  movel([0.274819, -1.341479, -2.579880, -0.791030, 1.570796, 1.845616],accel_mss,speed_ms,0,blend_radius_m)
  movel([0.275794, -1.341271, -2.580017, -0.791101, 1.570796, 1.846590],accel_mss,speed_ms,0,blend_radius_m)
  movel([0.276766, -1.341079, -2.580143, -0.791167, 1.570796, 1.847563],accel_mss,speed_ms,0,blend_radius_m)
  movel([0.277679, -1.340913, -2.580252, -0.791224, 1.570796, 1.848475],accel_mss,speed_ms,0,blend_radius_m)
  movel([0.278587, -1.340762, -2.580351, -0.791276, 1.570796, 1.849384],accel_mss,speed_ms,0,blend_radius_m)
  movel([0.278988, -1.340706, -2.580387, -0.791295, 1.570796, 1.849784],accel_mss,speed_ms,0,blend_radius_m)
  movel([0.279382, -1.340663, -2.580416, -0.791310, 1.570796, 1.850178],accel_mss,speed_ms,0,blend_radius_m)
  movel([0.279771, -1.340637, -2.580433, -0.791319, 1.570796, 1.850568],accel_mss,speed_ms,0,blend_radius_m)
  movel([0.279984, -1.340628, -2.580439, -0.791322, 1.570796, 1.850780],accel_mss,speed_ms,0,blend_radius_m)
  movel([0.280191, -1.340629, -2.580438, -0.791322, 1.570796, 1.850987],accel_mss,speed_ms,0,blend_radius_m)
  movel([0.280203, -1.340637, -2.580433, -0.791319, 1.570796, 1.850999],accel_mss,speed_ms,0,blend_radius_m)
  movel([0.280197, -1.340656, -2.580421, -0.791313, 1.570796, 1.850993],accel_mss,speed_ms,0,blend_radius_m)
  movel([0.280179, -1.340667, -2.580413, -0.791309, 1.570796, 1.850976],accel_mss,speed_ms,0,blend_radius_m)
  speed_ms = 0.003
  movel([0.280179, -1.327920, -2.574072, -0.810397, 1.570796, 1.850976],accel_mss,speed_ms,0,blend_radius_m)
  speed_ms = 0.01
  movel([0.280179, -1.303552, -2.561012, -0.847825, 1.570796, 1.850976],accel_mss,speed_ms,0,blend_radius_m)
  movel([0.262380, -1.358037, -2.525199, -0.829153, 1.570796, 1.833176],accel_mss,speed_ms,0,blend_radius_m)
  movel([0.262380, -1.381577, -2.537576, -0.793236, 1.570796, 1.833176],accel_mss,speed_ms,0,blend_radius_m)
  speed_ms = 0.003
  movel([0.262380, -1.390744, -2.542086, -0.779559, 1.570796, 1.833176],accel_mss,speed_ms,0,blend_radius_m)
  speed_ms = 0.007
  movel([0.261890, -1.392448, -2.540846, -0.779096, 1.570796, 1.832686],accel_mss,speed_ms,0,blend_radius_m)
  movel([0.261638, -1.393307, -2.540218, -0.778864, 1.570796, 1.832434],accel_mss,speed_ms,0,blend_radius_m)
  movel([0.261560, -1.393546, -2.540044, -0.778799, 1.570796, 1.832357],accel_mss,speed_ms,0,blend_radius_m)
  movel([0.261476, -1.393785, -2.539869, -0.778735, 1.570796, 1.832272],accel_mss,speed_ms,0,blend_radius_m)
  movel([0.261419, -1.393927, -2.539765, -0.778697, 1.570796, 1.832216],accel_mss,speed_ms,0,blend_radius_m)
  movel([0.261357, -1.394067, -2.539663, -0.778659, 1.570796, 1.832153],accel_mss,speed_ms,0,blend_radius_m)
  movel([0.261341, -1.394090, -2.539646, -0.778653, 1.570796, 1.832137],accel_mss,speed_ms,0,blend_radius_m)
  movel([0.261318, -1.394107, -2.539633, -0.778648, 1.570796, 1.832114],accel_mss,speed_ms,0,blend_radius_m)
  movel([0.261293, -1.394115, -2.539628, -0.778646, 1.570796, 1.832090],accel_mss,speed_ms,0,blend_radius_m)
  movel([0.261271, -1.394116, -2.539627, -0.778646, 1.570796, 1.832067],accel_mss,speed_ms,0,blend_radius_m)
  movel([0.256001, -1.393339, -2.540195, -0.778855, 1.570796, 1.826797],accel_mss,speed_ms,0,blend_radius_m)
  movel([0.256257, -1.392428, -2.540860, -0.779101, 1.570796, 1.827054],accel_mss,speed_ms,0,blend_radius_m)
  movel([0.256515, -1.391516, -2.541524, -0.779349, 1.570796, 1.827311],accel_mss,speed_ms,0,blend_radius_m)
  movel([0.259448, -1.391126, -2.541808, -0.779455, 1.570796, 1.830244],accel_mss,speed_ms,0,blend_radius_m)
  movel([0.262380, -1.390744, -2.542086, -0.779559, 1.570796, 1.833176],accel_mss,speed_ms,0,blend_radius_m)
  speed_ms = 0.003
  movel([0.262380, -1.393840, -2.543573, -0.774975, 1.570796, 1.833176],accel_mss,speed_ms,0,blend_radius_m)
  speed_ms = 0.007
  movel([0.261890, -1.395540, -2.542330, -0.774519, 1.570796, 1.832686],accel_mss,speed_ms,0,blend_radius_m)
  movel([0.261638, -1.396398, -2.541701, -0.774290, 1.570796, 1.832434],accel_mss,speed_ms,0,blend_radius_m)
  movel([0.261560, -1.396636, -2.541527, -0.774227, 1.570796, 1.832357],accel_mss,speed_ms,0,blend_radius_m)
  movel([0.261476, -1.396875, -2.541351, -0.774163, 1.570796, 1.832272],accel_mss,speed_ms,0,blend_radius_m)
  movel([0.261419, -1.397016, -2.541248, -0.774126, 1.570796, 1.832216],accel_mss,speed_ms,0,blend_radius_m)
  movel([0.261357, -1.397155, -2.541145, -0.774089, 1.570796, 1.832153],accel_mss,speed_ms,0,blend_radius_m)
  movel([0.261341, -1.397178, -2.541128, -0.774083, 1.570796, 1.832137],accel_mss,speed_ms,0,blend_radius_m)
  movel([0.261318, -1.397196, -2.541115, -0.774078, 1.570796, 1.832114],accel_mss,speed_ms,0,blend_radius_m)
  movel([0.261293, -1.397203, -2.541110, -0.774076, 1.570796, 1.832090],accel_mss,speed_ms,0,blend_radius_m)
  movel([0.261271, -1.397204, -2.541109, -0.774076, 1.570796, 1.832067],accel_mss,speed_ms,0,blend_radius_m)
  movel([0.256001, -1.396429, -2.541678, -0.774282, 1.570796, 1.826797],accel_mss,speed_ms,0,blend_radius_m)
  movel([0.256257, -1.395521, -2.542344, -0.774524, 1.570796, 1.827054],accel_mss,speed_ms,0,blend_radius_m)
  movel([0.256515, -1.394611, -2.543010, -0.774768, 1.570796, 1.827311],accel_mss,speed_ms,0,blend_radius_m)
  movel([0.259448, -1.394222, -2.543295, -0.774872, 1.570796, 1.830244],accel_mss,speed_ms,0,blend_radius_m)
  movel([0.262380, -1.393840, -2.543573, -0.774975, 1.570796, 1.833176],accel_mss,speed_ms,0,blend_radius_m)
  speed_ms = 0.003
  movel([0.262380, -1.381577, -2.537576, -0.793236, 1.570796, 1.833176],accel_mss,speed_ms,0,blend_radius_m)
  speed_ms = 0.01
  movel([0.262380, -1.358037, -2.525199, -0.829153, 1.570796, 1.833176],accel_mss,speed_ms,0,blend_radius_m)
  movel([0.278975, -1.298309, -2.564258, -0.849822, 1.570796, 1.849771],accel_mss,speed_ms,0,blend_radius_m)
  movel([0.278975, -1.322751, -2.577384, -0.812254, 1.570796, 1.849771],accel_mss,speed_ms,0,blend_radius_m)
  speed_ms = 0.003
  movel([0.278975, -1.332307, -2.582178, -0.797904, 1.570796, 1.849771],accel_mss,speed_ms,0,blend_radius_m)
  speed_ms = 0.007
  movel([0.275846, -1.332753, -2.581889, -0.797747, 1.570796, 1.846643],accel_mss,speed_ms,0,blend_radius_m)
  movel([0.272717, -1.333207, -2.581595, -0.797586, 1.570796, 1.843513],accel_mss,speed_ms,0,blend_radius_m)
  movel([0.273170, -1.331664, -2.582593, -0.798132, 1.570796, 1.843966],accel_mss,speed_ms,0,blend_radius_m)
  movel([0.273625, -1.330114, -2.583591, -0.798683, 1.570796, 1.844422],accel_mss,speed_ms,0,blend_radius_m)
  movel([0.274406, -1.330222, -2.583522, -0.798645, 1.570796, 1.845202],accel_mss,speed_ms,0,blend_radius_m)
  movel([0.274838, -1.330281, -2.583484, -0.798624, 1.570796, 1.845634],accel_mss,speed_ms,0,blend_radius_m)
  movel([0.275574, -1.330385, -2.583417, -0.798587, 1.570796, 1.846370],accel_mss,speed_ms,0,blend_radius_m)
  movel([0.276428, -1.330502, -2.583342, -0.798545, 1.570796, 1.847224],accel_mss,speed_ms,0,blend_radius_m)
  movel([0.277289, -1.330626, -2.583262, -0.798501, 1.570796, 1.848086],accel_mss,speed_ms,0,blend_radius_m)
  movel([0.279389, -1.330926, -2.583069, -0.798394, 1.570796, 1.850186],accel_mss,speed_ms,0,blend_radius_m)
  movel([0.279182, -1.331618, -2.582623, -0.798149, 1.570796, 1.849978],accel_mss,speed_ms,0,blend_radius_m)
  movel([0.278975, -1.332307, -2.582178, -0.797904, 1.570796, 1.849771],accel_mss,speed_ms,0,blend_radius_m)
  speed_ms = 0.003
  movel([0.278975, -1.335541, -2.583759, -0.793089, 1.570796, 1.849771],accel_mss,speed_ms,0,blend_radius_m)
  speed_ms = 0.007
  movel([0.275846, -1.335986, -2.583470, -0.792933, 1.570796, 1.846643],accel_mss,speed_ms,0,blend_radius_m)
  movel([0.272717, -1.336439, -2.583175, -0.792775, 1.570796, 1.843513],accel_mss,speed_ms,0,blend_radius_m)
  movel([0.273170, -1.334899, -2.584176, -0.793315, 1.570796, 1.843966],accel_mss,speed_ms,0,blend_radius_m)
  movel([0.273625, -1.333353, -2.585176, -0.793860, 1.570796, 1.844422],accel_mss,speed_ms,0,blend_radius_m)
  movel([0.274406, -1.333460, -2.585107, -0.793822, 1.570796, 1.845202],accel_mss,speed_ms,0,blend_radius_m)
  movel([0.274838, -1.333519, -2.585069, -0.793801, 1.570796, 1.845634],accel_mss,speed_ms,0,blend_radius_m)
  movel([0.275574, -1.333622, -2.585002, -0.793765, 1.570796, 1.846370],accel_mss,speed_ms,0,blend_radius_m)
  movel([0.276428, -1.333739, -2.584926, -0.793723, 1.570796, 1.847224],accel_mss,speed_ms,0,blend_radius_m)
  movel([0.277289, -1.333863, -2.584846, -0.793680, 1.570796, 1.848086],accel_mss,speed_ms,0,blend_radius_m)
  movel([0.279389, -1.334162, -2.584653, -0.793574, 1.570796, 1.850186],accel_mss,speed_ms,0,blend_radius_m)
  movel([0.279182, -1.334853, -2.584205, -0.793331, 1.570796, 1.849978],accel_mss,speed_ms,0,blend_radius_m)
  movel([0.278975, -1.335541, -2.583759, -0.793089, 1.570796, 1.849771],accel_mss,speed_ms,0,blend_radius_m)
  speed_ms = 0.003
  movel([0.278975, -1.322751, -2.577384, -0.812254, 1.570796, 1.849771],accel_mss,speed_ms,0,blend_radius_m)
  speed_ms = 0.01
  movel([0.278975, -1.298309, -2.564258, -0.849822, 1.570796, 1.849771],accel_mss,speed_ms,0,blend_radius_m)
  movel([0.264711, -1.307973, -2.558248, -0.846168, 1.570796, 1.835507],accel_mss,speed_ms,0,blend_radius_m)
  movel([0.264711, -1.332279, -2.571252, -0.808858, 1.570796, 1.835507],accel_mss,speed_ms,0,blend_radius_m)
  speed_ms = 0.003
  movel([0.264711, -1.341777, -2.575999, -0.794614, 1.570796, 1.835507],accel_mss,speed_ms,0,blend_radius_m)
  speed_ms = 0.007
  movel([0.264715, -1.341787, -2.575992, -0.794610, 1.570796, 1.835511],accel_mss,speed_ms,0,blend_radius_m)
  movel([0.264709, -1.341799, -2.575984, -0.794606, 1.570796, 1.835505],accel_mss,speed_ms,0,blend_radius_m)
  movel([0.264688, -1.341820, -2.575970, -0.794599, 1.570796, 1.835485],accel_mss,speed_ms,0,blend_radius_m)
  movel([0.264666, -1.341839, -2.575957, -0.794592, 1.570796, 1.835463],accel_mss,speed_ms,0,blend_radius_m)
  movel([0.264589, -1.341894, -2.575921, -0.794574, 1.570796, 1.835385],accel_mss,speed_ms,0,blend_radius_m)
  movel([0.264497, -1.341950, -2.575884, -0.794555, 1.570796, 1.835293],accel_mss,speed_ms,0,blend_radius_m)
  movel([0.264400, -1.341999, -2.575852, -0.794538, 1.570796, 1.835196],accel_mss,speed_ms,0,blend_radius_m)
  movel([0.264310, -1.342037, -2.575827, -0.794525, 1.570796, 1.835107],accel_mss,speed_ms,0,blend_radius_m)
  movel([0.264246, -1.342053, -2.575816, -0.794520, 1.570796, 1.835043],accel_mss,speed_ms,0,blend_radius_m)
  movel([0.264232, -1.342053, -2.575816, -0.794520, 1.570796, 1.835028],accel_mss,speed_ms,0,blend_radius_m)
  movel([0.264222, -1.342048, -2.575820, -0.794521, 1.570796, 1.835018],accel_mss,speed_ms,0,blend_radius_m)
  movel([0.264217, -1.342037, -2.575827, -0.794525, 1.570796, 1.835014],accel_mss,speed_ms,0,blend_radius_m)
  movel([0.264223, -1.342025, -2.575835, -0.794529, 1.570796, 1.835020],accel_mss,speed_ms,0,blend_radius_m)
  movel([0.264244, -1.342004, -2.575849, -0.794536, 1.570796, 1.835040],accel_mss,speed_ms,0,blend_radius_m)
  movel([0.264266, -1.341985, -2.575861, -0.794543, 1.570796, 1.835062],accel_mss,speed_ms,0,blend_radius_m)
  movel([0.264341, -1.341931, -2.575897, -0.794561, 1.570796, 1.835137],accel_mss,speed_ms,0,blend_radius_m)
  movel([0.264435, -1.341874, -2.575934, -0.794581, 1.570796, 1.835232],accel_mss,speed_ms,0,blend_radius_m)
  movel([0.264532, -1.341826, -2.575966, -0.794597, 1.570796, 1.835329],accel_mss,speed_ms,0,blend_radius_m)
  movel([0.264622, -1.341788, -2.575991, -0.794610, 1.570796, 1.835418],accel_mss,speed_ms,0,blend_radius_m)
  movel([0.264683, -1.341772, -2.576002, -0.794616, 1.570796, 1.835480],accel_mss,speed_ms,0,blend_radius_m)
  movel([0.264700, -1.341771, -2.576002, -0.794616, 1.570796, 1.835496],accel_mss,speed_ms,0,blend_radius_m)
  movel([0.264711, -1.341777, -2.575999, -0.794614, 1.570796, 1.835507],accel_mss,speed_ms,0,blend_radius_m)
  speed_ms = 0.003
  movel([0.264711, -1.344989, -2.577565, -0.789835, 1.570796, 1.835507],accel_mss,speed_ms,0,blend_radius_m)
  speed_ms = 0.007
  movel([0.264715, -1.345000, -2.577558, -0.789832, 1.570796, 1.835511],accel_mss,speed_ms,0,blend_radius_m)
  movel([0.264709, -1.345012, -2.577550, -0.789827, 1.570796, 1.835505],accel_mss,speed_ms,0,blend_radius_m)
  movel([0.264688, -1.345033, -2.577536, -0.789820, 1.570796, 1.835485],accel_mss,speed_ms,0,blend_radius_m)
  movel([0.264666, -1.345052, -2.577523, -0.789814, 1.570796, 1.835463],accel_mss,speed_ms,0,blend_radius_m)
  movel([0.264589, -1.345106, -2.577487, -0.789796, 1.570796, 1.835385],accel_mss,speed_ms,0,blend_radius_m)
  movel([0.264497, -1.345163, -2.577450, -0.789777, 1.570796, 1.835293],accel_mss,speed_ms,0,blend_radius_m)
  movel([0.264400, -1.345211, -2.577418, -0.789760, 1.570796, 1.835196],accel_mss,speed_ms,0,blend_radius_m)
  movel([0.264310, -1.345249, -2.577393, -0.789747, 1.570796, 1.835107],accel_mss,speed_ms,0,blend_radius_m)
  movel([0.264246, -1.345265, -2.577382, -0.789742, 1.570796, 1.835043],accel_mss,speed_ms,0,blend_radius_m)
  movel([0.264232, -1.345265, -2.577382, -0.789742, 1.570796, 1.835028],accel_mss,speed_ms,0,blend_radius_m)
  movel([0.264222, -1.345260, -2.577385, -0.789744, 1.570796, 1.835018],accel_mss,speed_ms,0,blend_radius_m)
  movel([0.264217, -1.345249, -2.577392, -0.789747, 1.570796, 1.835014],accel_mss,speed_ms,0,blend_radius_m)
  movel([0.264223, -1.345237, -2.577400, -0.789751, 1.570796, 1.835020],accel_mss,speed_ms,0,blend_radius_m)
  movel([0.264244, -1.345216, -2.577414, -0.789758, 1.570796, 1.835040],accel_mss,speed_ms,0,blend_radius_m)
  movel([0.264266, -1.345197, -2.577427, -0.789765, 1.570796, 1.835062],accel_mss,speed_ms,0,blend_radius_m)
  movel([0.264341, -1.345143, -2.577463, -0.789783, 1.570796, 1.835137],accel_mss,speed_ms,0,blend_radius_m)
  movel([0.264435, -1.345086, -2.577500, -0.789802, 1.570796, 1.835232],accel_mss,speed_ms,0,blend_radius_m)
  movel([0.264532, -1.345038, -2.577532, -0.789819, 1.570796, 1.835329],accel_mss,speed_ms,0,blend_radius_m)
  movel([0.264622, -1.345000, -2.577557, -0.789831, 1.570796, 1.835418],accel_mss,speed_ms,0,blend_radius_m)
  movel([0.264683, -1.344984, -2.577568, -0.789837, 1.570796, 1.835480],accel_mss,speed_ms,0,blend_radius_m)
  movel([0.264700, -1.344984, -2.577568, -0.789837, 1.570796, 1.835496],accel_mss,speed_ms,0,blend_radius_m)
  movel([0.264711, -1.344989, -2.577565, -0.789835, 1.570796, 1.835507],accel_mss,speed_ms,0,blend_radius_m)
  speed_ms = 0.003
  movel([0.264711, -1.332279, -2.571252, -0.808858, 1.570796, 1.835507],accel_mss,speed_ms,0,blend_radius_m)
  speed_ms = 0.01
  movel([0.264711, -1.307973, -2.558248, -0.846168, 1.570796, 1.835507],accel_mss,speed_ms,0,blend_radius_m)
  movel([0.264022, -1.308308, -2.558037, -0.846043, 1.570796, 1.834819],accel_mss,speed_ms,0,blend_radius_m)
  movel([0.264022, -1.332610, -2.571037, -0.808742, 1.570796, 1.834819],accel_mss,speed_ms,0,blend_radius_m)
  speed_ms = 0.003
  movel([0.264022, -1.342105, -2.575782, -0.794502, 1.570796, 1.834819],accel_mss,speed_ms,0,blend_radius_m)
  speed_ms = 0.007
  movel([0.264026, -1.342115, -2.575775, -0.794498, 1.570796, 1.834823],accel_mss,speed_ms,0,blend_radius_m)
  movel([0.264020, -1.342128, -2.575767, -0.794494, 1.570796, 1.834817],accel_mss,speed_ms,0,blend_radius_m)
  movel([0.264000, -1.342149, -2.575753, -0.794487, 1.570796, 1.834797],accel_mss,speed_ms,0,blend_radius_m)
  movel([0.263978, -1.342168, -2.575741, -0.794481, 1.570796, 1.834774],accel_mss,speed_ms,0,blend_radius_m)
  movel([0.263901, -1.342222, -2.575705, -0.794462, 1.570796, 1.834697],accel_mss,speed_ms,0,blend_radius_m)
  movel([0.263809, -1.342279, -2.575668, -0.794443, 1.570796, 1.834605],accel_mss,speed_ms,0,blend_radius_m)
  movel([0.263712, -1.342327, -2.575636, -0.794426, 1.570796, 1.834508],accel_mss,speed_ms,0,blend_radius_m)
  movel([0.263622, -1.342365, -2.575610, -0.794413, 1.570796, 1.834419],accel_mss,speed_ms,0,blend_radius_m)
  movel([0.263558, -1.342382, -2.575600, -0.794408, 1.570796, 1.834354],accel_mss,speed_ms,0,blend_radius_m)
  movel([0.263544, -1.342381, -2.575600, -0.794408, 1.570796, 1.834340],accel_mss,speed_ms,0,blend_radius_m)
  movel([0.263534, -1.342376, -2.575603, -0.794410, 1.570796, 1.834330],accel_mss,speed_ms,0,blend_radius_m)
  movel([0.263529, -1.342366, -2.575610, -0.794413, 1.570796, 1.834326],accel_mss,speed_ms,0,blend_radius_m)
  movel([0.263535, -1.342354, -2.575618, -0.794417, 1.570796, 1.834332],accel_mss,speed_ms,0,blend_radius_m)
  movel([0.263555, -1.342332, -2.575632, -0.794424, 1.570796, 1.834352],accel_mss,speed_ms,0,blend_radius_m)
  movel([0.263578, -1.342313, -2.575645, -0.794431, 1.570796, 1.834374],accel_mss,speed_ms,0,blend_radius_m)
  movel([0.263652, -1.342259, -2.575680, -0.794449, 1.570796, 1.834449],accel_mss,speed_ms,0,blend_radius_m)
  movel([0.263747, -1.342202, -2.575718, -0.794469, 1.570796, 1.834543],accel_mss,speed_ms,0,blend_radius_m)
  movel([0.263844, -1.342154, -2.575750, -0.794485, 1.570796, 1.834640],accel_mss,speed_ms,0,blend_radius_m)
  movel([0.263933, -1.342116, -2.575775, -0.794498, 1.570796, 1.834730],accel_mss,speed_ms,0,blend_radius_m)
  movel([0.263995, -1.342100, -2.575785, -0.794504, 1.570796, 1.834791],accel_mss,speed_ms,0,blend_radius_m)
  movel([0.264012, -1.342100, -2.575786, -0.794504, 1.570796, 1.834808],accel_mss,speed_ms,0,blend_radius_m)
  movel([0.264022, -1.342105, -2.575782, -0.794502, 1.570796, 1.834819],accel_mss,speed_ms,0,blend_radius_m)
  speed_ms = 0.003
  movel([0.264022, -1.345317, -2.577348, -0.789725, 1.570796, 1.834819],accel_mss,speed_ms,0,blend_radius_m)
  speed_ms = 0.007
  movel([0.264026, -1.345327, -2.577341, -0.789721, 1.570796, 1.834823],accel_mss,speed_ms,0,blend_radius_m)
  movel([0.264020, -1.345339, -2.577333, -0.789717, 1.570796, 1.834817],accel_mss,speed_ms,0,blend_radius_m)
  movel([0.264000, -1.345360, -2.577319, -0.789710, 1.570796, 1.834797],accel_mss,speed_ms,0,blend_radius_m)
  movel([0.263978, -1.345379, -2.577306, -0.789703, 1.570796, 1.834774],accel_mss,speed_ms,0,blend_radius_m)
  movel([0.263901, -1.345434, -2.577270, -0.789685, 1.570796, 1.834697],accel_mss,speed_ms,0,blend_radius_m)
  movel([0.263809, -1.345490, -2.577233, -0.789666, 1.570796, 1.834605],accel_mss,speed_ms,0,blend_radius_m)
  movel([0.263712, -1.345538, -2.577201, -0.789650, 1.570796, 1.834508],accel_mss,speed_ms,0,blend_radius_m)
  movel([0.263622, -1.345576, -2.577176, -0.789637, 1.570796, 1.834419],accel_mss,speed_ms,0,blend_radius_m)
  movel([0.263558, -1.345593, -2.577165, -0.789631, 1.570796, 1.834354],accel_mss,speed_ms,0,blend_radius_m)
  movel([0.263544, -1.345593, -2.577165, -0.789631, 1.570796, 1.834340],accel_mss,speed_ms,0,blend_radius_m)
  movel([0.263534, -1.345588, -2.577168, -0.789633, 1.570796, 1.834330],accel_mss,speed_ms,0,blend_radius_m)
  movel([0.263529, -1.345577, -2.577175, -0.789637, 1.570796, 1.834326],accel_mss,speed_ms,0,blend_radius_m)
  movel([0.263535, -1.345565, -2.577183, -0.789641, 1.570796, 1.834332],accel_mss,speed_ms,0,blend_radius_m)
  movel([0.263555, -1.345544, -2.577197, -0.789648, 1.570796, 1.834352],accel_mss,speed_ms,0,blend_radius_m)
  movel([0.263578, -1.345525, -2.577210, -0.789654, 1.570796, 1.834374],accel_mss,speed_ms,0,blend_radius_m)
  movel([0.263652, -1.345471, -2.577246, -0.789672, 1.570796, 1.834449],accel_mss,speed_ms,0,blend_radius_m)
  movel([0.263747, -1.345414, -2.577283, -0.789692, 1.570796, 1.834543],accel_mss,speed_ms,0,blend_radius_m)
  movel([0.263844, -1.345366, -2.577315, -0.789708, 1.570796, 1.834640],accel_mss,speed_ms,0,blend_radius_m)
  movel([0.263933, -1.345328, -2.577340, -0.789721, 1.570796, 1.834730],accel_mss,speed_ms,0,blend_radius_m)
  movel([0.263995, -1.345312, -2.577351, -0.789726, 1.570796, 1.834791],accel_mss,speed_ms,0,blend_radius_m)
  movel([0.264012, -1.345311, -2.577351, -0.789726, 1.570796, 1.834808],accel_mss,speed_ms,0,blend_radius_m)
  movel([0.264022, -1.345317, -2.577348, -0.789725, 1.570796, 1.834819],accel_mss,speed_ms,0,blend_radius_m)
  speed_ms = 0.003
  movel([0.264022, -1.332610, -2.571037, -0.808742, 1.570796, 1.834819],accel_mss,speed_ms,0,blend_radius_m)
  speed_ms = 0.01
  movel([0.264022, -1.308308, -2.558037, -0.846043, 1.570796, 1.834819],accel_mss,speed_ms,0,blend_radius_m)
  movel([0.248737, -1.294338, -2.566693, -0.851357, 1.570796, 1.819533],accel_mss,speed_ms,0,blend_radius_m)
  movel([0.248737, -1.318834, -2.579871, -0.813685, 1.570796, 1.819533],accel_mss,speed_ms,0,blend_radius_m)
  speed_ms = 0.003
  movel([0.248737, -1.328414, -2.584683, -0.799292, 1.570796, 1.819533],accel_mss,speed_ms,0,blend_radius_m)
  speed_ms = 0.007
  movel([0.248697, -1.328446, -2.584662, -0.799280, 1.570796, 1.819493],accel_mss,speed_ms,0,blend_radius_m)
  movel([0.248652, -1.328468, -2.584649, -0.799273, 1.570796, 1.819448],accel_mss,speed_ms,0,blend_radius_m)
  movel([0.245500, -1.329570, -2.583941, -0.798878, 1.570796, 1.816296],accel_mss,speed_ms,0,blend_radius_m)
  movel([0.242434, -1.330648, -2.583248, -0.798493, 1.570796, 1.813230],accel_mss,speed_ms,0,blend_radius_m)
  movel([0.242300, -1.330689, -2.583221, -0.798479, 1.570796, 1.813096],accel_mss,speed_ms,0,blend_radius_m)
  movel([0.242169, -1.330719, -2.583202, -0.798468, 1.570796, 1.812965],accel_mss,speed_ms,0,blend_radius_m)
  movel([0.242113, -1.330722, -2.583200, -0.798467, 1.570796, 1.812909],accel_mss,speed_ms,0,blend_radius_m)
  movel([0.242059, -1.330716, -2.583204, -0.798469, 1.570796, 1.812855],accel_mss,speed_ms,0,blend_radius_m)
  movel([0.240657, -1.330365, -2.583430, -0.798594, 1.570796, 1.811454],accel_mss,speed_ms,0,blend_radius_m)
  movel([0.239079, -1.329963, -2.583689, -0.798737, 1.570796, 1.809875],accel_mss,speed_ms,0,blend_radius_m)
  movel([0.237230, -1.329485, -2.583996, -0.798908, 1.570796, 1.808027],accel_mss,speed_ms,0,blend_radius_m)
  movel([0.231703, -1.328086, -2.584894, -0.799410, 1.570796, 1.802500],accel_mss,speed_ms,0,blend_radius_m)
  movel([0.232587, -1.326228, -2.586081, -0.800080, 1.570796, 1.803383],accel_mss,speed_ms,0,blend_radius_m)
  movel([0.232933, -1.325504, -2.586543, -0.800342, 1.570796, 1.803729],accel_mss,speed_ms,0,blend_radius_m)
  movel([0.233237, -1.324867, -2.586949, -0.800574, 1.570796, 1.804034],accel_mss,speed_ms,0,blend_radius_m)
  movel([0.233502, -1.324323, -2.587294, -0.800772, 1.570796, 1.804298],accel_mss,speed_ms,0,blend_radius_m)
  movel([0.233562, -1.324211, -2.587365, -0.800812, 1.570796, 1.804358],accel_mss,speed_ms,0,blend_radius_m)
  movel([0.233589, -1.324181, -2.587385, -0.800823, 1.570796, 1.804385],accel_mss,speed_ms,0,blend_radius_m)
  movel([0.233622, -1.324163, -2.587396, -0.800830, 1.570796, 1.804419],accel_mss,speed_ms,0,blend_radius_m)
  movel([0.233654, -1.324164, -2.587395, -0.800829, 1.570796, 1.804450],accel_mss,speed_ms,0,blend_radius_m)
  movel([0.234609, -1.324536, -2.587159, -0.800694, 1.570796, 1.805405],accel_mss,speed_ms,0,blend_radius_m)
  movel([0.235192, -1.324772, -2.587009, -0.800608, 1.570796, 1.805988],accel_mss,speed_ms,0,blend_radius_m)
  movel([0.235770, -1.325013, -2.586855, -0.800520, 1.570796, 1.806567],accel_mss,speed_ms,0,blend_radius_m)
  movel([0.236518, -1.325343, -2.586646, -0.800401, 1.570796, 1.807314],accel_mss,speed_ms,0,blend_radius_m)
  movel([0.237265, -1.325673, -2.586435, -0.800281, 1.570796, 1.808061],accel_mss,speed_ms,0,blend_radius_m)
  movel([0.239935, -1.326833, -2.585695, -0.799861, 1.570796, 1.810731],accel_mss,speed_ms,0,blend_radius_m)
  movel([0.240884, -1.327196, -2.585463, -0.799730, 1.570796, 1.811680],accel_mss,speed_ms,0,blend_radius_m)
  movel([0.240920, -1.327178, -2.585474, -0.799737, 1.570796, 1.811716],accel_mss,speed_ms,0,blend_radius_m)
  movel([0.240947, -1.327148, -2.585493, -0.799747, 1.570796, 1.811743],accel_mss,speed_ms,0,blend_radius_m)
  movel([0.244595, -1.319268, -2.590491, -0.802631, 1.570796, 1.815391],accel_mss,speed_ms,0,blend_radius_m)
  movel([0.245457, -1.317406, -2.591659, -0.803324, 1.570796, 1.816253],accel_mss,speed_ms,0,blend_radius_m)
  movel([0.246216, -1.315769, -2.592683, -0.803937, 1.570796, 1.817013],accel_mss,speed_ms,0,blend_radius_m)
  movel([0.246297, -1.315594, -2.592792, -0.804003, 1.570796, 1.817093],accel_mss,speed_ms,0,blend_radius_m)
  movel([0.246319, -1.315390, -2.592920, -0.804079, 1.570796, 1.817115],accel_mss,speed_ms,0,blend_radius_m)
  movel([0.239012, -1.318049, -2.591256, -0.803084, 1.570796, 1.809808],accel_mss,speed_ms,0,blend_radius_m)
  movel([0.237328, -1.318654, -2.590876, -0.802859, 1.570796, 1.808124],accel_mss,speed_ms,0,blend_radius_m)
  movel([0.235834, -1.319181, -2.590545, -0.802663, 1.570796, 1.806630],accel_mss,speed_ms,0,blend_radius_m)
  movel([0.235811, -1.319185, -2.590542, -0.802661, 1.570796, 1.806607],accel_mss,speed_ms,0,blend_radius_m)
  movel([0.235795, -1.319179, -2.590546, -0.802664, 1.570796, 1.806592],accel_mss,speed_ms,0,blend_radius_m)
  movel([0.235787, -1.319162, -2.590557, -0.802670, 1.570796, 1.806584],accel_mss,speed_ms,0,blend_radius_m)
  movel([0.235786, -1.319121, -2.590583, -0.802685, 1.570796, 1.806582],accel_mss,speed_ms,0,blend_radius_m)
  movel([0.235792, -1.319076, -2.590611, -0.802702, 1.570796, 1.806589],accel_mss,speed_ms,0,blend_radius_m)
  movel([0.235811, -1.319031, -2.590640, -0.802719, 1.570796, 1.806607],accel_mss,speed_ms,0,blend_radius_m)
  movel([0.236634, -1.317353, -2.591693, -0.803344, 1.570796, 1.807431],accel_mss,speed_ms,0,blend_radius_m)
  movel([0.237464, -1.315667, -2.592747, -0.803975, 1.570796, 1.808260],accel_mss,speed_ms,0,blend_radius_m)
  movel([0.237489, -1.315625, -2.592773, -0.803991, 1.570796, 1.808285],accel_mss,speed_ms,0,blend_radius_m)
  movel([0.237524, -1.315587, -2.592797, -0.804005, 1.570796, 1.808320],accel_mss,speed_ms,0,blend_radius_m)
  movel([0.237562, -1.315552, -2.592819, -0.804019, 1.570796, 1.808358],accel_mss,speed_ms,0,blend_radius_m)
  movel([0.237608, -1.315527, -2.592834, -0.804028, 1.570796, 1.808404],accel_mss,speed_ms,0,blend_radius_m)
  movel([0.239936, -1.314636, -2.593389, -0.804363, 1.570796, 1.810732],accel_mss,speed_ms,0,blend_radius_m)
  movel([0.242517, -1.313656, -2.594000, -0.804734, 1.570796, 1.813313],accel_mss,speed_ms,0,blend_radius_m)
  movel([0.245578, -1.312504, -2.594715, -0.805170, 1.570796, 1.816374],accel_mss,speed_ms,0,blend_radius_m)
  movel([0.253566, -1.309525, -2.596557, -0.806308, 1.570796, 1.824362],accel_mss,speed_ms,0,blend_radius_m)
  movel([0.255227, -1.311268, -2.595480, -0.805641, 1.570796, 1.826023],accel_mss,speed_ms,0,blend_radius_m)
  movel([0.255862, -1.311938, -2.595065, -0.805385, 1.570796, 1.826658],accel_mss,speed_ms,0,blend_radius_m)
  movel([0.256392, -1.312512, -2.594710, -0.805167, 1.570796, 1.827189],accel_mss,speed_ms,0,blend_radius_m)
  movel([0.256867, -1.313027, -2.594390, -0.804972, 1.570796, 1.827663],accel_mss,speed_ms,0,blend_radius_m)
  movel([0.256871, -1.313038, -2.594383, -0.804968, 1.570796, 1.827667],accel_mss,speed_ms,0,blend_radius_m)
  movel([0.256869, -1.313055, -2.594373, -0.804961, 1.570796, 1.827665],accel_mss,speed_ms,0,blend_radius_m)
  movel([0.256857, -1.313087, -2.594353, -0.804949, 1.570796, 1.827654],accel_mss,speed_ms,0,blend_radius_m)
  movel([0.255658, -1.315350, -2.592944, -0.804094, 1.570796, 1.826455],accel_mss,speed_ms,0,blend_radius_m)
  movel([0.254339, -1.317843, -2.591385, -0.803161, 1.570796, 1.825135],accel_mss,speed_ms,0,blend_radius_m)
  movel([0.252782, -1.320784, -2.589536, -0.802070, 1.570796, 1.823579],accel_mss,speed_ms,0,blend_radius_m)
  movel([0.251233, -1.323711, -2.587683, -0.800995, 1.570796, 1.822029],accel_mss,speed_ms,0,blend_radius_m)
  movel([0.249932, -1.326169, -2.586119, -0.800101, 1.570796, 1.820728],accel_mss,speed_ms,0,blend_radius_m)
  movel([0.248759, -1.328385, -2.584701, -0.799302, 1.570796, 1.819555],accel_mss,speed_ms,0,blend_radius_m)
  movel([0.248737, -1.328414, -2.584683, -0.799292, 1.570796, 1.819533],accel_mss,speed_ms,0,blend_radius_m)
  speed_ms = 0.003
  movel([0.248737, -1.331656, -2.586271, -0.794462, 1.570796, 1.819533],accel_mss,speed_ms,0,blend_radius_m)
  speed_ms = 0.007
  movel([0.248697, -1.331688, -2.586250, -0.794450, 1.570796, 1.819493],accel_mss,speed_ms,0,blend_radius_m)
  movel([0.248652, -1.331709, -2.586237, -0.794443, 1.570796, 1.819448],accel_mss,speed_ms,0,blend_radius_m)
  movel([0.245500, -1.332810, -2.585527, -0.794052, 1.570796, 1.816296],accel_mss,speed_ms,0,blend_radius_m)
  movel([0.242434, -1.333885, -2.584832, -0.793672, 1.570796, 1.813230],accel_mss,speed_ms,0,blend_radius_m)
  movel([0.242300, -1.333926, -2.584806, -0.793657, 1.570796, 1.813096],accel_mss,speed_ms,0,blend_radius_m)
  movel([0.242169, -1.333956, -2.584786, -0.793647, 1.570796, 1.812965],accel_mss,speed_ms,0,blend_radius_m)
  movel([0.242113, -1.333959, -2.584784, -0.793646, 1.570796, 1.812909],accel_mss,speed_ms,0,blend_radius_m)
  movel([0.242059, -1.333953, -2.584788, -0.793648, 1.570796, 1.812855],accel_mss,speed_ms,0,blend_radius_m)
  movel([0.240657, -1.333602, -2.585015, -0.793772, 1.570796, 1.811454],accel_mss,speed_ms,0,blend_radius_m)
  movel([0.239079, -1.333201, -2.585274, -0.793913, 1.570796, 1.809875],accel_mss,speed_ms,0,blend_radius_m)
  movel([0.237230, -1.332725, -2.585582, -0.794082, 1.570796, 1.808027],accel_mss,speed_ms,0,blend_radius_m)
  movel([0.231703, -1.331328, -2.586482, -0.794579, 1.570796, 1.802500],accel_mss,speed_ms,0,blend_radius_m)
  movel([0.232587, -1.329475, -2.587673, -0.795242, 1.570796, 1.803383],accel_mss,speed_ms,0,blend_radius_m)
  movel([0.232933, -1.328752, -2.588136, -0.795501, 1.570796, 1.803729],accel_mss,speed_ms,0,blend_radius_m)
  movel([0.233237, -1.328116, -2.588543, -0.795730, 1.570796, 1.804034],accel_mss,speed_ms,0,blend_radius_m)
  movel([0.233502, -1.327574, -2.588889, -0.795926, 1.570796, 1.804298],accel_mss,speed_ms,0,blend_radius_m)
  movel([0.233562, -1.327462, -2.588960, -0.795966, 1.570796, 1.804358],accel_mss,speed_ms,0,blend_radius_m)
  movel([0.233589, -1.327432, -2.588979, -0.795977, 1.570796, 1.804385],accel_mss,speed_ms,0,blend_radius_m)
  movel([0.233622, -1.327415, -2.588991, -0.795984, 1.570796, 1.804419],accel_mss,speed_ms,0,blend_radius_m)
  movel([0.233654, -1.327416, -2.588990, -0.795983, 1.570796, 1.804450],accel_mss,speed_ms,0,blend_radius_m)
  movel([0.234609, -1.327787, -2.588753, -0.795849, 1.570796, 1.805405],accel_mss,speed_ms,0,blend_radius_m)
  movel([0.235192, -1.328022, -2.588603, -0.795764, 1.570796, 1.805988],accel_mss,speed_ms,0,blend_radius_m)
  movel([0.235770, -1.328262, -2.588449, -0.795678, 1.570796, 1.806567],accel_mss,speed_ms,0,blend_radius_m)
  movel([0.236518, -1.328591, -2.588239, -0.795559, 1.570796, 1.807314],accel_mss,speed_ms,0,blend_radius_m)
  movel([0.237265, -1.328921, -2.588028, -0.795441, 1.570796, 1.808061],accel_mss,speed_ms,0,blend_radius_m)
  movel([0.239935, -1.330079, -2.587285, -0.795025, 1.570796, 1.810731],accel_mss,speed_ms,0,blend_radius_m)
  movel([0.240884, -1.330441, -2.587053, -0.794896, 1.570796, 1.811680],accel_mss,speed_ms,0,blend_radius_m)
  movel([0.240920, -1.330423, -2.587064, -0.794902, 1.570796, 1.811716],accel_mss,speed_ms,0,blend_radius_m)
  movel([0.240947, -1.330393, -2.587084, -0.794913, 1.570796, 1.811743],accel_mss,speed_ms,0,blend_radius_m)
  movel([0.244595, -1.322529, -2.592094, -0.797766, 1.570796, 1.815391],accel_mss,speed_ms,0,blend_radius_m)
  movel([0.245457, -1.320671, -2.593265, -0.798452, 1.570796, 1.816253],accel_mss,speed_ms,0,blend_radius_m)
  movel([0.246216, -1.319038, -2.594292, -0.799059, 1.570796, 1.817013],accel_mss,speed_ms,0,blend_radius_m)
  movel([0.246297, -1.318863, -2.594401, -0.799124, 1.570796, 1.817093],accel_mss,speed_ms,0,blend_radius_m)
  movel([0.246319, -1.318660, -2.594529, -0.799200, 1.570796, 1.817115],accel_mss,speed_ms,0,blend_radius_m)
  movel([0.239012, -1.321313, -2.592861, -0.798215, 1.570796, 1.809808],accel_mss,speed_ms,0,blend_radius_m)
  movel([0.237328, -1.321917, -2.592480, -0.797992, 1.570796, 1.808124],accel_mss,speed_ms,0,blend_radius_m)
  movel([0.235834, -1.322443, -2.592148, -0.797798, 1.570796, 1.806630],accel_mss,speed_ms,0,blend_radius_m)
  movel([0.235811, -1.322447, -2.592146, -0.797796, 1.570796, 1.806607],accel_mss,speed_ms,0,blend_radius_m)
  movel([0.235795, -1.322441, -2.592149, -0.797799, 1.570796, 1.806592],accel_mss,speed_ms,0,blend_radius_m)
  movel([0.235787, -1.322424, -2.592160, -0.797805, 1.570796, 1.806584],accel_mss,speed_ms,0,blend_radius_m)
  movel([0.235786, -1.322383, -2.592186, -0.797820, 1.570796, 1.806582],accel_mss,speed_ms,0,blend_radius_m)
  movel([0.235792, -1.322338, -2.592215, -0.797837, 1.570796, 1.806589],accel_mss,speed_ms,0,blend_radius_m)
  movel([0.235811, -1.322293, -2.592243, -0.797853, 1.570796, 1.806607],accel_mss,speed_ms,0,blend_radius_m)
  movel([0.236634, -1.320618, -2.593299, -0.798472, 1.570796, 1.807431],accel_mss,speed_ms,0,blend_radius_m)
  movel([0.237464, -1.318936, -2.594356, -0.799097, 1.570796, 1.808260],accel_mss,speed_ms,0,blend_radius_m)
  movel([0.237489, -1.318895, -2.594382, -0.799113, 1.570796, 1.808285],accel_mss,speed_ms,0,blend_radius_m)
  movel([0.237524, -1.318856, -2.594406, -0.799127, 1.570796, 1.808320],accel_mss,speed_ms,0,blend_radius_m)
  movel([0.237562, -1.318821, -2.594428, -0.799140, 1.570796, 1.808358],accel_mss,speed_ms,0,blend_radius_m)
  movel([0.237608, -1.318796, -2.594443, -0.799149, 1.570796, 1.808404],accel_mss,speed_ms,0,blend_radius_m)
  movel([0.239936, -1.317908, -2.595000, -0.799481, 1.570796, 1.810732],accel_mss,speed_ms,0,blend_radius_m)
  movel([0.242517, -1.316929, -2.595612, -0.799848, 1.570796, 1.813313],accel_mss,speed_ms,0,blend_radius_m)
  movel([0.245578, -1.315779, -2.596329, -0.800281, 1.570796, 1.816374],accel_mss,speed_ms,0,blend_radius_m)
  movel([0.253566, -1.312806, -2.598176, -0.801407, 1.570796, 1.824362],accel_mss,speed_ms,0,blend_radius_m)
  movel([0.255227, -1.314546, -2.597096, -0.800746, 1.570796, 1.826023],accel_mss,speed_ms,0,blend_radius_m)
  movel([0.255862, -1.315215, -2.596680, -0.800493, 1.570796, 1.826658],accel_mss,speed_ms,0,blend_radius_m)
  movel([0.256392, -1.315788, -2.596324, -0.800277, 1.570796, 1.827189],accel_mss,speed_ms,0,blend_radius_m)
  movel([0.256867, -1.316302, -2.596003, -0.800084, 1.570796, 1.827663],accel_mss,speed_ms,0,blend_radius_m)
  movel([0.256871, -1.316313, -2.595997, -0.800080, 1.570796, 1.827667],accel_mss,speed_ms,0,blend_radius_m)
  movel([0.256869, -1.316329, -2.595986, -0.800073, 1.570796, 1.827665],accel_mss,speed_ms,0,blend_radius_m)
  movel([0.256857, -1.316362, -2.595966, -0.800061, 1.570796, 1.827654],accel_mss,speed_ms,0,blend_radius_m)
  movel([0.255658, -1.318620, -2.594554, -0.799215, 1.570796, 1.826455],accel_mss,speed_ms,0,blend_radius_m)
  movel([0.254339, -1.321108, -2.592991, -0.798291, 1.570796, 1.825135],accel_mss,speed_ms,0,blend_radius_m)
  movel([0.252782, -1.324042, -2.591136, -0.797211, 1.570796, 1.823579],accel_mss,speed_ms,0,blend_radius_m)
  movel([0.251233, -1.326963, -2.589279, -0.796147, 1.570796, 1.822029],accel_mss,speed_ms,0,blend_radius_m)
  movel([0.249932, -1.329416, -2.587710, -0.795263, 1.570796, 1.820728],accel_mss,speed_ms,0,blend_radius_m)
  movel([0.248759, -1.331627, -2.586289, -0.794472, 1.570796, 1.819555],accel_mss,speed_ms,0,blend_radius_m)
  movel([0.248737, -1.331656, -2.586271, -0.794462, 1.570796, 1.819533],accel_mss,speed_ms,0,blend_radius_m)
  speed_ms = 0.003
  movel([0.248737, -1.318834, -2.579871, -0.813685, 1.570796, 1.819533],accel_mss,speed_ms,0,blend_radius_m)
  speed_ms = 0.01
  movel([0.248737, -1.294338, -2.566693, -0.851357, 1.570796, 1.819533],accel_mss,speed_ms,0,blend_radius_m)
  movel([0.235155, -1.310004, -2.556970, -0.845415, 1.570796, 1.805951],accel_mss,speed_ms,0,blend_radius_m)
  movel([0.235155, -1.334281, -2.569948, -0.808160, 1.570796, 1.805951],accel_mss,speed_ms,0,blend_radius_m)
  speed_ms = 0.003
  movel([0.235155, -1.343766, -2.574685, -0.793938, 1.570796, 1.805951],accel_mss,speed_ms,0,blend_radius_m)
  speed_ms = 0.007
  movel([0.234636, -1.345662, -2.573428, -0.793299, 1.570796, 1.805432],accel_mss,speed_ms,0,blend_radius_m)
  movel([0.234118, -1.347555, -2.572169, -0.792665, 1.570796, 1.804915],accel_mss,speed_ms,0,blend_radius_m)
  movel([0.226584, -1.353832, -2.567957, -0.790600, 1.570796, 1.797380],accel_mss,speed_ms,0,blend_radius_m)
  movel([0.219134, -1.360071, -2.563718, -0.788601, 1.570796, 1.789930],accel_mss,speed_ms,0,blend_radius_m)
  movel([0.218563, -1.362440, -2.562093, -0.787856, 1.570796, 1.789359],accel_mss,speed_ms,0,blend_radius_m)
  movel([0.217996, -1.364798, -2.560469, -0.787122, 1.570796, 1.788792],accel_mss,speed_ms,0,blend_radius_m)
  movel([0.214308, -1.365470, -2.560005, -0.786914, 1.570796, 1.785105],accel_mss,speed_ms,0,blend_radius_m)
  movel([0.212898, -1.365727, -2.559827, -0.786835, 1.570796, 1.783694],accel_mss,speed_ms,0,blend_radius_m)
  movel([0.211722, -1.365934, -2.559684, -0.786771, 1.570796, 1.782518],accel_mss,speed_ms,0,blend_radius_m)
  movel([0.210685, -1.366114, -2.559560, -0.786716, 1.570796, 1.781482],accel_mss,speed_ms,0,blend_radius_m)
  movel([0.210677, -1.366109, -2.559563, -0.786717, 1.570796, 1.781473],accel_mss,speed_ms,0,blend_radius_m)
  movel([0.210682, -1.366097, -2.559571, -0.786721, 1.570796, 1.781479],accel_mss,speed_ms,0,blend_radius_m)
  movel([0.210705, -1.366078, -2.559585, -0.786727, 1.570796, 1.781502],accel_mss,speed_ms,0,blend_radius_m)
  movel([0.210733, -1.366062, -2.559596, -0.786731, 1.570796, 1.781529],accel_mss,speed_ms,0,blend_radius_m)
  movel([0.211085, -1.365874, -2.559726, -0.786789, 1.570796, 1.781882],accel_mss,speed_ms,0,blend_radius_m)
  movel([0.211496, -1.365660, -2.559874, -0.786855, 1.570796, 1.782292],accel_mss,speed_ms,0,blend_radius_m)
  movel([0.211972, -1.365414, -2.560044, -0.786931, 1.570796, 1.782768],accel_mss,speed_ms,0,blend_radius_m)
  movel([0.213200, -1.364790, -2.560475, -0.787124, 1.570796, 1.783996],accel_mss,speed_ms,0,blend_radius_m)
  movel([0.213474, -1.363625, -2.561278, -0.787486, 1.570796, 1.784271],accel_mss,speed_ms,0,blend_radius_m)
  movel([0.213749, -1.362459, -2.562080, -0.787850, 1.570796, 1.784545],accel_mss,speed_ms,0,blend_radius_m)
  movel([0.215855, -1.361496, -2.562741, -0.788151, 1.570796, 1.786651],accel_mss,speed_ms,0,blend_radius_m)
  movel([0.217964, -1.360535, -2.563399, -0.788454, 1.570796, 1.788761],accel_mss,speed_ms,0,blend_radius_m)
  movel([0.219239, -1.355234, -2.567009, -0.790146, 1.570796, 1.790035],accel_mss,speed_ms,0,blend_radius_m)
  movel([0.220529, -1.349889, -2.570609, -0.791891, 1.570796, 1.791325],accel_mss,speed_ms,0,blend_radius_m)
  movel([0.218685, -1.349648, -2.570770, -0.791971, 1.570796, 1.789481],accel_mss,speed_ms,0,blend_radius_m)
  movel([0.216839, -1.349412, -2.570928, -0.792049, 1.570796, 1.787635],accel_mss,speed_ms,0,blend_radius_m)
  movel([0.217085, -1.348375, -2.571621, -0.792392, 1.570796, 1.787882],accel_mss,speed_ms,0,blend_radius_m)
  movel([0.217333, -1.347338, -2.572314, -0.792738, 1.570796, 1.788129],accel_mss,speed_ms,0,blend_radius_m)
  movel([0.216967, -1.347252, -2.572370, -0.792766, 1.570796, 1.787763],accel_mss,speed_ms,0,blend_radius_m)
  movel([0.216949, -1.347238, -2.572380, -0.792771, 1.570796, 1.787745],accel_mss,speed_ms,0,blend_radius_m)
  movel([0.216944, -1.347217, -2.572394, -0.792778, 1.570796, 1.787740],accel_mss,speed_ms,0,blend_radius_m)
  movel([0.216955, -1.347190, -2.572412, -0.792787, 1.570796, 1.787751],accel_mss,speed_ms,0,blend_radius_m)
  movel([0.216980, -1.347166, -2.572428, -0.792795, 1.570796, 1.787776],accel_mss,speed_ms,0,blend_radius_m)
  movel([0.217007, -1.347154, -2.572436, -0.792799, 1.570796, 1.787803],accel_mss,speed_ms,0,blend_radius_m)
  movel([0.217637, -1.347010, -2.572532, -0.792847, 1.570796, 1.788434],accel_mss,speed_ms,0,blend_radius_m)
  movel([0.218263, -1.346876, -2.572621, -0.792892, 1.570796, 1.789059],accel_mss,speed_ms,0,blend_radius_m)
  movel([0.219422, -1.346641, -2.572778, -0.792971, 1.570796, 1.790218],accel_mss,speed_ms,0,blend_radius_m)
  movel([0.220577, -1.346417, -2.572926, -0.793045, 1.570796, 1.791374],accel_mss,speed_ms,0,blend_radius_m)
  movel([0.225877, -1.345431, -2.573582, -0.793376, 1.570796, 1.796674],accel_mss,speed_ms,0,blend_radius_m)
  movel([0.235155, -1.343766, -2.574685, -0.793938, 1.570796, 1.805951],accel_mss,speed_ms,0,blend_radius_m)
  speed_ms = 0.003
  movel([0.235155, -1.346974, -2.576248, -0.789167, 1.570796, 1.805951],accel_mss,speed_ms,0,blend_radius_m)
  speed_ms = 0.007
  movel([0.234636, -1.348866, -2.574988, -0.788535, 1.570796, 1.805432],accel_mss,speed_ms,0,blend_radius_m)
  movel([0.234118, -1.350754, -2.573725, -0.787909, 1.570796, 1.804915],accel_mss,speed_ms,0,blend_radius_m)
  movel([0.226584, -1.357017, -2.569504, -0.785868, 1.570796, 1.797380],accel_mss,speed_ms,0,blend_radius_m)
  movel([0.219134, -1.363241, -2.565254, -0.783894, 1.570796, 1.789930],accel_mss,speed_ms,0,blend_radius_m)
  movel([0.218563, -1.365605, -2.563626, -0.783158, 1.570796, 1.789359],accel_mss,speed_ms,0,blend_radius_m)
  movel([0.217996, -1.367958, -2.561998, -0.782433, 1.570796, 1.788792],accel_mss,speed_ms,0,blend_radius_m)
  movel([0.214308, -1.368628, -2.561533, -0.782228, 1.570796, 1.785105],accel_mss,speed_ms,0,blend_radius_m)
  movel([0.212898, -1.368884, -2.561355, -0.782150, 1.570796, 1.783694],accel_mss,speed_ms,0,blend_radius_m)
  movel([0.211722, -1.369091, -2.561211, -0.782087, 1.570796, 1.782518],accel_mss,speed_ms,0,blend_radius_m)
  movel([0.210685, -1.369270, -2.561086, -0.782032, 1.570796, 1.781482],accel_mss,speed_ms,0,blend_radius_m)
  movel([0.210677, -1.369265, -2.561090, -0.782034, 1.570796, 1.781473],accel_mss,speed_ms,0,blend_radius_m)
  movel([0.210682, -1.369254, -2.561098, -0.782037, 1.570796, 1.781479],accel_mss,speed_ms,0,blend_radius_m)
  movel([0.210705, -1.369234, -2.561111, -0.782043, 1.570796, 1.781502],accel_mss,speed_ms,0,blend_radius_m)
  movel([0.210733, -1.369218, -2.561122, -0.782048, 1.570796, 1.781529],accel_mss,speed_ms,0,blend_radius_m)
  movel([0.211085, -1.369031, -2.561253, -0.782105, 1.570796, 1.781882],accel_mss,speed_ms,0,blend_radius_m)
  movel([0.211496, -1.368817, -2.561401, -0.782170, 1.570796, 1.782292],accel_mss,speed_ms,0,blend_radius_m)
  movel([0.211972, -1.368572, -2.561572, -0.782245, 1.570796, 1.782768],accel_mss,speed_ms,0,blend_radius_m)
  movel([0.213200, -1.367950, -2.562003, -0.782436, 1.570796, 1.783996],accel_mss,speed_ms,0,blend_radius_m)
  movel([0.213474, -1.366787, -2.562809, -0.782793, 1.570796, 1.784271],accel_mss,speed_ms,0,blend_radius_m)
  movel([0.213749, -1.365624, -2.563613, -0.783152, 1.570796, 1.784545],accel_mss,speed_ms,0,blend_radius_m)
  movel([0.215855, -1.364664, -2.564275, -0.783450, 1.570796, 1.786651],accel_mss,speed_ms,0,blend_radius_m)
  movel([0.217964, -1.363705, -2.564935, -0.783749, 1.570796, 1.788761],accel_mss,speed_ms,0,blend_radius_m)
  movel([0.219239, -1.358416, -2.568553, -0.785420, 1.570796, 1.790035],accel_mss,speed_ms,0,blend_radius_m)
  movel([0.220529, -1.353083, -2.572162, -0.787144, 1.570796, 1.791325],accel_mss,speed_ms,0,blend_radius_m)
  movel([0.218685, -1.352843, -2.572323, -0.787222, 1.570796, 1.789481],accel_mss,speed_ms,0,blend_radius_m)
  movel([0.216839, -1.352607, -2.572482, -0.787300, 1.570796, 1.787635],accel_mss,speed_ms,0,blend_radius_m)
  movel([0.217085, -1.351573, -2.573177, -0.787639, 1.570796, 1.787882],accel_mss,speed_ms,0,blend_radius_m)
  movel([0.217333, -1.350538, -2.573871, -0.787981, 1.570796, 1.788129],accel_mss,speed_ms,0,blend_radius_m)
  movel([0.216967, -1.350452, -2.573928, -0.788009, 1.570796, 1.787763],accel_mss,speed_ms,0,blend_radius_m)
  movel([0.216949, -1.350438, -2.573937, -0.788014, 1.570796, 1.787745],accel_mss,speed_ms,0,blend_radius_m)
  movel([0.216944, -1.350417, -2.573951, -0.788021, 1.570796, 1.787740],accel_mss,speed_ms,0,blend_radius_m)
  movel([0.216955, -1.350391, -2.573969, -0.788029, 1.570796, 1.787751],accel_mss,speed_ms,0,blend_radius_m)
  movel([0.216980, -1.350366, -2.573985, -0.788037, 1.570796, 1.787776],accel_mss,speed_ms,0,blend_radius_m)
  movel([0.217007, -1.350355, -2.573993, -0.788041, 1.570796, 1.787803],accel_mss,speed_ms,0,blend_radius_m)
  movel([0.217637, -1.350211, -2.574089, -0.788089, 1.570796, 1.788434],accel_mss,speed_ms,0,blend_radius_m)
  movel([0.218263, -1.350078, -2.574179, -0.788133, 1.570796, 1.789059],accel_mss,speed_ms,0,blend_radius_m)
  movel([0.219422, -1.349842, -2.574336, -0.788211, 1.570796, 1.790218],accel_mss,speed_ms,0,blend_radius_m)
  movel([0.220577, -1.349619, -2.574485, -0.788285, 1.570796, 1.791374],accel_mss,speed_ms,0,blend_radius_m)
  movel([0.225877, -1.348635, -2.575142, -0.788612, 1.570796, 1.796674],accel_mss,speed_ms,0,blend_radius_m)
  movel([0.235155, -1.346974, -2.576248, -0.789167, 1.570796, 1.805951],accel_mss,speed_ms,0,blend_radius_m)
  speed_ms = 0.003
  movel([0.235155, -1.334281, -2.569948, -0.808160, 1.570796, 1.805951],accel_mss,speed_ms,0,blend_radius_m)
  speed_ms = 0.01
  movel([0.235155, -1.310004, -2.556970, -0.845415, 1.570796, 1.805951],accel_mss,speed_ms,0,blend_radius_m)
  movel([0.233548, -1.315976, -2.553182, -0.843231, 1.570796, 1.804344],accel_mss,speed_ms,0,blend_radius_m)
  movel([0.233548, -1.340167, -2.566085, -0.806138, 1.570796, 1.804344],accel_mss,speed_ms,0,blend_radius_m)
  speed_ms = 0.003
  movel([0.233548, -1.349613, -2.570793, -0.791982, 1.570796, 1.804344],accel_mss,speed_ms,0,blend_radius_m)
  speed_ms = 0.007
  movel([0.233570, -1.349609, -2.570796, -0.791983, 1.570796, 1.804366],accel_mss,speed_ms,0,blend_radius_m)
  movel([0.233584, -1.349618, -2.570790, -0.791981, 1.570796, 1.804381],accel_mss,speed_ms,0,blend_radius_m)
  movel([0.233587, -1.349635, -2.570779, -0.791975, 1.570796, 1.804383],accel_mss,speed_ms,0,blend_radius_m)
  movel([0.233141, -1.351503, -2.569526, -0.791360, 1.570796, 1.803938],accel_mss,speed_ms,0,blend_radius_m)
  movel([0.232881, -1.352579, -2.568802, -0.791008, 1.570796, 1.803678],accel_mss,speed_ms,0,blend_radius_m)
  movel([0.232615, -1.353652, -2.568079, -0.790659, 1.570796, 1.803412],accel_mss,speed_ms,0,blend_radius_m)
  movel([0.231949, -1.356298, -2.566288, -0.789803, 1.570796, 1.802746],accel_mss,speed_ms,0,blend_radius_m)
  movel([0.230259, -1.362970, -2.561729, -0.787690, 1.570796, 1.801055],accel_mss,speed_ms,0,blend_radius_m)
  movel([0.226624, -1.363595, -2.561299, -0.787495, 1.570796, 1.797421],accel_mss,speed_ms,0,blend_radius_m)
  movel([0.225106, -1.363853, -2.561121, -0.787415, 1.570796, 1.795902],accel_mss,speed_ms,0,blend_radius_m)
  movel([0.223550, -1.364111, -2.560943, -0.787335, 1.570796, 1.794346],accel_mss,speed_ms,0,blend_radius_m)
  movel([0.222167, -1.364333, -2.560790, -0.787266, 1.570796, 1.792963],accel_mss,speed_ms,0,blend_radius_m)
  movel([0.221716, -1.364400, -2.560744, -0.787245, 1.570796, 1.792512],accel_mss,speed_ms,0,blend_radius_m)
  movel([0.221265, -1.364465, -2.560699, -0.787225, 1.570796, 1.792061],accel_mss,speed_ms,0,blend_radius_m)
  movel([0.219540, -1.364702, -2.560536, -0.787151, 1.570796, 1.790336],accel_mss,speed_ms,0,blend_radius_m)
  movel([0.220062, -1.362544, -2.562022, -0.787823, 1.570796, 1.790858],accel_mss,speed_ms,0,blend_radius_m)
  movel([0.220587, -1.360376, -2.563508, -0.788504, 1.570796, 1.791384],accel_mss,speed_ms,0,blend_radius_m)
  movel([0.226976, -1.355038, -2.567142, -0.790209, 1.570796, 1.797773],accel_mss,speed_ms,0,blend_radius_m)
  movel([0.229452, -1.352979, -2.568532, -0.790877, 1.570796, 1.800248],accel_mss,speed_ms,0,blend_radius_m)
  movel([0.231562, -1.351233, -2.569707, -0.791449, 1.570796, 1.802359],accel_mss,speed_ms,0,blend_radius_m)
  movel([0.233456, -1.349673, -2.570753, -0.791962, 1.570796, 1.804253],accel_mss,speed_ms,0,blend_radius_m)
  movel([0.233500, -1.349642, -2.570775, -0.791973, 1.570796, 1.804296],accel_mss,speed_ms,0,blend_radius_m)
  movel([0.233548, -1.349613, -2.570793, -0.791982, 1.570796, 1.804344],accel_mss,speed_ms,0,blend_radius_m)
  speed_ms = 0.003
  movel([0.233548, -1.352808, -2.572347, -0.787234, 1.570796, 1.804344],accel_mss,speed_ms,0,blend_radius_m)
  speed_ms = 0.007
  movel([0.233570, -1.352804, -2.572349, -0.787235, 1.570796, 1.804366],accel_mss,speed_ms,0,blend_radius_m)
  movel([0.233584, -1.352813, -2.572344, -0.787232, 1.570796, 1.804381],accel_mss,speed_ms,0,blend_radius_m)
  movel([0.233587, -1.352830, -2.572332, -0.787227, 1.570796, 1.804383],accel_mss,speed_ms,0,blend_radius_m)
  movel([0.233141, -1.354693, -2.571076, -0.786619, 1.570796, 1.803938],accel_mss,speed_ms,0,blend_radius_m)
  movel([0.232881, -1.355767, -2.570351, -0.786272, 1.570796, 1.803678],accel_mss,speed_ms,0,blend_radius_m)
  movel([0.232615, -1.356837, -2.569625, -0.785926, 1.570796, 1.803412],accel_mss,speed_ms,0,blend_radius_m)
  movel([0.231949, -1.359478, -2.567830, -0.785081, 1.570796, 1.802746],accel_mss,speed_ms,0,blend_radius_m)
  movel([0.230259, -1.366134, -2.563261, -0.782994, 1.570796, 1.801055],accel_mss,speed_ms,0,blend_radius_m)
  movel([0.226624, -1.366758, -2.562829, -0.782802, 1.570796, 1.797421],accel_mss,speed_ms,0,blend_radius_m)
  movel([0.225106, -1.367015, -2.562651, -0.782723, 1.570796, 1.795902],accel_mss,speed_ms,0,blend_radius_m)
  movel([0.223550, -1.367272, -2.562473, -0.782644, 1.570796, 1.794346],accel_mss,speed_ms,0,blend_radius_m)
  movel([0.222167, -1.367494, -2.562320, -0.782575, 1.570796, 1.792963],accel_mss,speed_ms,0,blend_radius_m)
  movel([0.221716, -1.367561, -2.562273, -0.782555, 1.570796, 1.792512],accel_mss,speed_ms,0,blend_radius_m)
  movel([0.221265, -1.367626, -2.562228, -0.782535, 1.570796, 1.792061],accel_mss,speed_ms,0,blend_radius_m)
  movel([0.219540, -1.367862, -2.562065, -0.782463, 1.570796, 1.790336],accel_mss,speed_ms,0,blend_radius_m)
  movel([0.220062, -1.365709, -2.563554, -0.783126, 1.570796, 1.790858],accel_mss,speed_ms,0,blend_radius_m)
  movel([0.220587, -1.363546, -2.565044, -0.783798, 1.570796, 1.791384],accel_mss,speed_ms,0,blend_radius_m)
  movel([0.226976, -1.358220, -2.568686, -0.785482, 1.570796, 1.797773],accel_mss,speed_ms,0,blend_radius_m)
  movel([0.229452, -1.356166, -2.570080, -0.786142, 1.570796, 1.800248],accel_mss,speed_ms,0,blend_radius_m)
  movel([0.231562, -1.354424, -2.571258, -0.786707, 1.570796, 1.802359],accel_mss,speed_ms,0,blend_radius_m)
  movel([0.233456, -1.352868, -2.572307, -0.787214, 1.570796, 1.804253],accel_mss,speed_ms,0,blend_radius_m)
  movel([0.233500, -1.352836, -2.572328, -0.787225, 1.570796, 1.804296],accel_mss,speed_ms,0,blend_radius_m)
  movel([0.233548, -1.352808, -2.572347, -0.787234, 1.570796, 1.804344],accel_mss,speed_ms,0,blend_radius_m)
  speed_ms = 0.003
  movel([0.233548, -1.340167, -2.566085, -0.806138, 1.570796, 1.804344],accel_mss,speed_ms,0,blend_radius_m)
  speed_ms = 0.01
  movel([0.233548, -1.315976, -2.553182, -0.843231, 1.570796, 1.804344],accel_mss,speed_ms,0,blend_radius_m)
  movel([0.227152, -1.342252, -2.535972, -0.834165, 1.570796, 1.797948],accel_mss,speed_ms,0,blend_radius_m)
  movel([0.227152, -1.366045, -2.548544, -0.797800, 1.570796, 1.797948],accel_mss,speed_ms,0,blend_radius_m)
  speed_ms = 0.003
  movel([0.227152, -1.375319, -2.553129, -0.783941, 1.570796, 1.797948],accel_mss,speed_ms,0,blend_radius_m)
  speed_ms = 0.007
  movel([0.225532, -1.381803, -2.548528, -0.782058, 1.570796, 1.796328],accel_mss,speed_ms,0,blend_radius_m)
  movel([0.224876, -1.384410, -2.546661, -0.781318, 1.570796, 1.795673],accel_mss,speed_ms,0,blend_radius_m)
  movel([0.224617, -1.385426, -2.545931, -0.781032, 1.570796, 1.795413],accel_mss,speed_ms,0,blend_radius_m)
  movel([0.224351, -1.386442, -2.545199, -0.780747, 1.570796, 1.795147],accel_mss,speed_ms,0,blend_radius_m)
  movel([0.223893, -1.388169, -2.543953, -0.780267, 1.570796, 1.794689],accel_mss,speed_ms,0,blend_radius_m)
  movel([0.223881, -1.388190, -2.543938, -0.780261, 1.570796, 1.794677],accel_mss,speed_ms,0,blend_radius_m)
  movel([0.223859, -1.388204, -2.543927, -0.780257, 1.570796, 1.794655],accel_mss,speed_ms,0,blend_radius_m)
  movel([0.223838, -1.388208, -2.543925, -0.780256, 1.570796, 1.794634],accel_mss,speed_ms,0,blend_radius_m)
  movel([0.223802, -1.388195, -2.543934, -0.780260, 1.570796, 1.794599],accel_mss,speed_ms,0,blend_radius_m)
  movel([0.223770, -1.388177, -2.543947, -0.780265, 1.570796, 1.794566],accel_mss,speed_ms,0,blend_radius_m)
  movel([0.222568, -1.387209, -2.544646, -0.780533, 1.570796, 1.793365],accel_mss,speed_ms,0,blend_radius_m)
  movel([0.221223, -1.386126, -2.545427, -0.780836, 1.570796, 1.792019],accel_mss,speed_ms,0,blend_radius_m)
  movel([0.219640, -1.384844, -2.546349, -0.781195, 1.570796, 1.790437],accel_mss,speed_ms,0,blend_radius_m)
  movel([0.215501, -1.381512, -2.548736, -0.782141, 1.570796, 1.786297],accel_mss,speed_ms,0,blend_radius_m)
  movel([0.216005, -1.379403, -2.550238, -0.782748, 1.570796, 1.786801],accel_mss,speed_ms,0,blend_radius_m)
  movel([0.216511, -1.377288, -2.551738, -0.783363, 1.570796, 1.787307],accel_mss,speed_ms,0,blend_radius_m)
  movel([0.218717, -1.376832, -2.552061, -0.783497, 1.570796, 1.789513],accel_mss,speed_ms,0,blend_radius_m)
  movel([0.219782, -1.376619, -2.552211, -0.783559, 1.570796, 1.790579],accel_mss,speed_ms,0,blend_radius_m)
  movel([0.221190, -1.376354, -2.552398, -0.783637, 1.570796, 1.791987],accel_mss,speed_ms,0,blend_radius_m)
  movel([0.222684, -1.376080, -2.552592, -0.783717, 1.570796, 1.793481],accel_mss,speed_ms,0,blend_radius_m)
  movel([0.224038, -1.375845, -2.552758, -0.783786, 1.570796, 1.794834],accel_mss,speed_ms,0,blend_radius_m)
  movel([0.227152, -1.375319, -2.553129, -0.783941, 1.570796, 1.797948],accel_mss,speed_ms,0,blend_radius_m)
  speed_ms = 0.003
  movel([0.227152, -1.378454, -2.554640, -0.779295, 1.570796, 1.797948],accel_mss,speed_ms,0,blend_radius_m)
  speed_ms = 0.007
  movel([0.225532, -1.384922, -2.550029, -0.777438, 1.570796, 1.796328],accel_mss,speed_ms,0,blend_radius_m)
  movel([0.224876, -1.387522, -2.548159, -0.776708, 1.570796, 1.795673],accel_mss,speed_ms,0,blend_radius_m)
  movel([0.224617, -1.388536, -2.547427, -0.776426, 1.570796, 1.795413],accel_mss,speed_ms,0,blend_radius_m)
  movel([0.224351, -1.389550, -2.546693, -0.776146, 1.570796, 1.795147],accel_mss,speed_ms,0,blend_radius_m)
  movel([0.223893, -1.391272, -2.545444, -0.775673, 1.570796, 1.794689],accel_mss,speed_ms,0,blend_radius_m)
  movel([0.223881, -1.391293, -2.545429, -0.775667, 1.570796, 1.794677],accel_mss,speed_ms,0,blend_radius_m)
  movel([0.223859, -1.391307, -2.545419, -0.775663, 1.570796, 1.794655],accel_mss,speed_ms,0,blend_radius_m)
  movel([0.223838, -1.391311, -2.545416, -0.775662, 1.570796, 1.794634],accel_mss,speed_ms,0,blend_radius_m)
  movel([0.223802, -1.391298, -2.545426, -0.775666, 1.570796, 1.794599],accel_mss,speed_ms,0,blend_radius_m)
  movel([0.223770, -1.391280, -2.545439, -0.775670, 1.570796, 1.794566],accel_mss,speed_ms,0,blend_radius_m)
  movel([0.222568, -1.390315, -2.546139, -0.775935, 1.570796, 1.793365],accel_mss,speed_ms,0,blend_radius_m)
  movel([0.221223, -1.389234, -2.546922, -0.776233, 1.570796, 1.792019],accel_mss,speed_ms,0,blend_radius_m)
  movel([0.219640, -1.387956, -2.547846, -0.776587, 1.570796, 1.790437],accel_mss,speed_ms,0,blend_radius_m)
  movel([0.215501, -1.384631, -2.550238, -0.777520, 1.570796, 1.786297],accel_mss,speed_ms,0,blend_radius_m)
  movel([0.216005, -1.382528, -2.551743, -0.778118, 1.570796, 1.786801],accel_mss,speed_ms,0,blend_radius_m)
  movel([0.216511, -1.380418, -2.553247, -0.778724, 1.570796, 1.787307],accel_mss,speed_ms,0,blend_radius_m)
  movel([0.218717, -1.379963, -2.553570, -0.778856, 1.570796, 1.789513],accel_mss,speed_ms,0,blend_radius_m)
  movel([0.219782, -1.379750, -2.553721, -0.778918, 1.570796, 1.790579],accel_mss,speed_ms,0,blend_radius_m)
  movel([0.221190, -1.379486, -2.553909, -0.778994, 1.570796, 1.791987],accel_mss,speed_ms,0,blend_radius_m)
  movel([0.222684, -1.379213, -2.554102, -0.779074, 1.570796, 1.793481],accel_mss,speed_ms,0,blend_radius_m)
  movel([0.224038, -1.378978, -2.554269, -0.779142, 1.570796, 1.794834],accel_mss,speed_ms,0,blend_radius_m)
  movel([0.227152, -1.378454, -2.554640, -0.779295, 1.570796, 1.797948],accel_mss,speed_ms,0,blend_radius_m)
  speed_ms = 0.003
  movel([0.227152, -1.366045, -2.548544, -0.797800, 1.570796, 1.797948],accel_mss,speed_ms,0,blend_radius_m)
  speed_ms = 0.01
  movel([0.227152, -1.342252, -2.535972, -0.834165, 1.570796, 1.797948],accel_mss,speed_ms,0,blend_radius_m)
  movel([0.215084, -1.343947, -2.534831, -0.833611, 1.570796, 1.785881],accel_mss,speed_ms,0,blend_radius_m)
  movel([0.215084, -1.367713, -2.547382, -0.797294, 1.570796, 1.785881],accel_mss,speed_ms,0,blend_radius_m)
  speed_ms = 0.003
  movel([0.215084, -1.376976, -2.551959, -0.783454, 1.570796, 1.785881],accel_mss,speed_ms,0,blend_radius_m)
  speed_ms = 0.007
  movel([0.214443, -1.379674, -2.550045, -0.782670, 1.570796, 1.785239],accel_mss,speed_ms,0,blend_radius_m)
  movel([0.213806, -1.382361, -2.548129, -0.781899, 1.570796, 1.784602],accel_mss,speed_ms,0,blend_radius_m)
  movel([0.217775, -1.385536, -2.545852, -0.781001, 1.570796, 1.788572],accel_mss,speed_ms,0,blend_radius_m)
  movel([0.219350, -1.386809, -2.544935, -0.780645, 1.570796, 1.790147],accel_mss,speed_ms,0,blend_radius_m)
  movel([0.220811, -1.388003, -2.544073, -0.780313, 1.570796, 1.791608],accel_mss,speed_ms,0,blend_radius_m)
  movel([0.222037, -1.389007, -2.543346, -0.780036, 1.570796, 1.792833],accel_mss,speed_ms,0,blend_radius_m)
  movel([0.222579, -1.389459, -2.543019, -0.779911, 1.570796, 1.793375],accel_mss,speed_ms,0,blend_radius_m)
  movel([0.223448, -1.390194, -2.542485, -0.779709, 1.570796, 1.794244],accel_mss,speed_ms,0,blend_radius_m)
  movel([0.223223, -1.391105, -2.541823, -0.779460, 1.570796, 1.794019],accel_mss,speed_ms,0,blend_radius_m)
  movel([0.222998, -1.392015, -2.541161, -0.779213, 1.570796, 1.793794],accel_mss,speed_ms,0,blend_radius_m)
  movel([0.214751, -1.393392, -2.540156, -0.778841, 1.570796, 1.785547],accel_mss,speed_ms,0,blend_radius_m)
  movel([0.206501, -1.394825, -2.539108, -0.778456, 1.570796, 1.777297],accel_mss,speed_ms,0,blend_radius_m)
  movel([0.206806, -1.393654, -2.539965, -0.778770, 1.570796, 1.777603],accel_mss,speed_ms,0,blend_radius_m)
  movel([0.207110, -1.392484, -2.540819, -0.779086, 1.570796, 1.777907],accel_mss,speed_ms,0,blend_radius_m)
  movel([0.209133, -1.391578, -2.541479, -0.779332, 1.570796, 1.779930],accel_mss,speed_ms,0,blend_radius_m)
  movel([0.211159, -1.390674, -2.542137, -0.779578, 1.570796, 1.781955],accel_mss,speed_ms,0,blend_radius_m)
  movel([0.212318, -1.385833, -2.545638, -0.780918, 1.570796, 1.783114],accel_mss,speed_ms,0,blend_radius_m)
  movel([0.212767, -1.383957, -2.546986, -0.781446, 1.570796, 1.783564],accel_mss,speed_ms,0,blend_radius_m)
  movel([0.213158, -1.382341, -2.548143, -0.781905, 1.570796, 1.783954],accel_mss,speed_ms,0,blend_radius_m)
  movel([0.213503, -1.380919, -2.549159, -0.782311, 1.570796, 1.784300],accel_mss,speed_ms,0,blend_radius_m)
  movel([0.213540, -1.380776, -2.549261, -0.782353, 1.570796, 1.784336],accel_mss,speed_ms,0,blend_radius_m)
  movel([0.213539, -1.380710, -2.549307, -0.782371, 1.570796, 1.784335],accel_mss,speed_ms,0,blend_radius_m)
  movel([0.213498, -1.380671, -2.549335, -0.782383, 1.570796, 1.784294],accel_mss,speed_ms,0,blend_radius_m)
  movel([0.213200, -1.380576, -2.549403, -0.782410, 1.570796, 1.783996],accel_mss,speed_ms,0,blend_radius_m)
  movel([0.212688, -1.380473, -2.549476, -0.782439, 1.570796, 1.783484],accel_mss,speed_ms,0,blend_radius_m)
  movel([0.209966, -1.380096, -2.549745, -0.782548, 1.570796, 1.780763],accel_mss,speed_ms,0,blend_radius_m)
  movel([0.210192, -1.379127, -2.550434, -0.782828, 1.570796, 1.780988],accel_mss,speed_ms,0,blend_radius_m)
  movel([0.210348, -1.378291, -2.551027, -0.783071, 1.570796, 1.781144],accel_mss,speed_ms,0,blend_radius_m)
  movel([0.210336, -1.378211, -2.551084, -0.783094, 1.570796, 1.781133],accel_mss,speed_ms,0,blend_radius_m)
  movel([0.210304, -1.378140, -2.551134, -0.783114, 1.570796, 1.781100],accel_mss,speed_ms,0,blend_radius_m)
  movel([0.210188, -1.378032, -2.551211, -0.783146, 1.570796, 1.780985],accel_mss,speed_ms,0,blend_radius_m)
  movel([0.210174, -1.378016, -2.551222, -0.783151, 1.570796, 1.780970],accel_mss,speed_ms,0,blend_radius_m)
  movel([0.210172, -1.377993, -2.551239, -0.783157, 1.570796, 1.780969],accel_mss,speed_ms,0,blend_radius_m)
  movel([0.210185, -1.377967, -2.551257, -0.783165, 1.570796, 1.780981],accel_mss,speed_ms,0,blend_radius_m)
  movel([0.210207, -1.377944, -2.551273, -0.783172, 1.570796, 1.781003],accel_mss,speed_ms,0,blend_radius_m)
  movel([0.210264, -1.377904, -2.551301, -0.783183, 1.570796, 1.781061],accel_mss,speed_ms,0,blend_radius_m)
  movel([0.210327, -1.377874, -2.551323, -0.783192, 1.570796, 1.781123],accel_mss,speed_ms,0,blend_radius_m)
  movel([0.210387, -1.377855, -2.551337, -0.783198, 1.570796, 1.781183],accel_mss,speed_ms,0,blend_radius_m)
  movel([0.210673, -1.377786, -2.551385, -0.783218, 1.570796, 1.781470],accel_mss,speed_ms,0,blend_radius_m)
  movel([0.210957, -1.377728, -2.551426, -0.783235, 1.570796, 1.781753],accel_mss,speed_ms,0,blend_radius_m)
  movel([0.212521, -1.377440, -2.551630, -0.783319, 1.570796, 1.783318],accel_mss,speed_ms,0,blend_radius_m)
  movel([0.215084, -1.376976, -2.551959, -0.783454, 1.570796, 1.785881],accel_mss,speed_ms,0,blend_radius_m)
  speed_ms = 0.003
  movel([0.215084, -1.380107, -2.553468, -0.778814, 1.570796, 1.785881],accel_mss,speed_ms,0,blend_radius_m)
  speed_ms = 0.007
  movel([0.214443, -1.382798, -2.551550, -0.778041, 1.570796, 1.785239],accel_mss,speed_ms,0,blend_radius_m)
  movel([0.213806, -1.385479, -2.549629, -0.777281, 1.570796, 1.784602],accel_mss,speed_ms,0,blend_radius_m)
  movel([0.217775, -1.388646, -2.547348, -0.776396, 1.570796, 1.788572],accel_mss,speed_ms,0,blend_radius_m)
  movel([0.219350, -1.389915, -2.546429, -0.776045, 1.570796, 1.790147],accel_mss,speed_ms,0,blend_radius_m)
  movel([0.220811, -1.391106, -2.545565, -0.775718, 1.570796, 1.791608],accel_mss,speed_ms,0,blend_radius_m)
  movel([0.222037, -1.392108, -2.544836, -0.775444, 1.570796, 1.792833],accel_mss,speed_ms,0,blend_radius_m)
  movel([0.222579, -1.392559, -2.544508, -0.775322, 1.570796, 1.793375],accel_mss,speed_ms,0,blend_radius_m)
  movel([0.223448, -1.393293, -2.543973, -0.775123, 1.570796, 1.794244],accel_mss,speed_ms,0,blend_radius_m)
  movel([0.223223, -1.394201, -2.543310, -0.774878, 1.570796, 1.794019],accel_mss,speed_ms,0,blend_radius_m)
  movel([0.222998, -1.395109, -2.542646, -0.774634, 1.570796, 1.793794],accel_mss,speed_ms,0,blend_radius_m)
  movel([0.214751, -1.396483, -2.541639, -0.774267, 1.570796, 1.785547],accel_mss,speed_ms,0,blend_radius_m)
  movel([0.206501, -1.397912, -2.540589, -0.773889, 1.570796, 1.777297],accel_mss,speed_ms,0,blend_radius_m)
  movel([0.206806, -1.396744, -2.541447, -0.774198, 1.570796, 1.777603],accel_mss,speed_ms,0,blend_radius_m)
  movel([0.207110, -1.395576, -2.542304, -0.774509, 1.570796, 1.777907],accel_mss,speed_ms,0,blend_radius_m)
  movel([0.209133, -1.394673, -2.542965, -0.774751, 1.570796, 1.779930],accel_mss,speed_ms,0,blend_radius_m)
  movel([0.211159, -1.393771, -2.543624, -0.774994, 1.570796, 1.781955],accel_mss,speed_ms,0,blend_radius_m)
  movel([0.212318, -1.388942, -2.547133, -0.776314, 1.570796, 1.783114],accel_mss,speed_ms,0,blend_radius_m)
  movel([0.212767, -1.387071, -2.548484, -0.776834, 1.570796, 1.783564],accel_mss,speed_ms,0,blend_radius_m)
  movel([0.213158, -1.385458, -2.549644, -0.777286, 1.570796, 1.783954],accel_mss,speed_ms,0,blend_radius_m)
  movel([0.213503, -1.384040, -2.550662, -0.777687, 1.570796, 1.784300],accel_mss,speed_ms,0,blend_radius_m)
  movel([0.213540, -1.383897, -2.550764, -0.777728, 1.570796, 1.784336],accel_mss,speed_ms,0,blend_radius_m)
  movel([0.213539, -1.383832, -2.550811, -0.777747, 1.570796, 1.784335],accel_mss,speed_ms,0,blend_radius_m)
  movel([0.213498, -1.383793, -2.550839, -0.777758, 1.570796, 1.784294],accel_mss,speed_ms,0,blend_radius_m)
  movel([0.213200, -1.383698, -2.550906, -0.777785, 1.570796, 1.783996],accel_mss,speed_ms,0,blend_radius_m)
  movel([0.212688, -1.383595, -2.550980, -0.777814, 1.570796, 1.783484],accel_mss,speed_ms,0,blend_radius_m)
  movel([0.209966, -1.383219, -2.551249, -0.777921, 1.570796, 1.780763],accel_mss,speed_ms,0,blend_radius_m)
  movel([0.210192, -1.382252, -2.551940, -0.778197, 1.570796, 1.780988],accel_mss,speed_ms,0,blend_radius_m)
  movel([0.210348, -1.381419, -2.552534, -0.778436, 1.570796, 1.781144],accel_mss,speed_ms,0,blend_radius_m)
  movel([0.210336, -1.381338, -2.552591, -0.778459, 1.570796, 1.781133],accel_mss,speed_ms,0,blend_radius_m)
  movel([0.210304, -1.381268, -2.552641, -0.778479, 1.570796, 1.781100],accel_mss,speed_ms,0,blend_radius_m)
  movel([0.210188, -1.381160, -2.552718, -0.778510, 1.570796, 1.780985],accel_mss,speed_ms,0,blend_radius_m)
  movel([0.210174, -1.381144, -2.552730, -0.778515, 1.570796, 1.780970],accel_mss,speed_ms,0,blend_radius_m)
  movel([0.210172, -1.381121, -2.552746, -0.778522, 1.570796, 1.780969],accel_mss,speed_ms,0,blend_radius_m)
  movel([0.210185, -1.381096, -2.552764, -0.778529, 1.570796, 1.780981],accel_mss,speed_ms,0,blend_radius_m)
  movel([0.210207, -1.381073, -2.552781, -0.778536, 1.570796, 1.781003],accel_mss,speed_ms,0,blend_radius_m)
  movel([0.210264, -1.381033, -2.552809, -0.778547, 1.570796, 1.781061],accel_mss,speed_ms,0,blend_radius_m)
  movel([0.210327, -1.381002, -2.552831, -0.778556, 1.570796, 1.781123],accel_mss,speed_ms,0,blend_radius_m)
  movel([0.210387, -1.380983, -2.552844, -0.778561, 1.570796, 1.781183],accel_mss,speed_ms,0,blend_radius_m)
  movel([0.210673, -1.380914, -2.552893, -0.778581, 1.570796, 1.781470],accel_mss,speed_ms,0,blend_radius_m)
  movel([0.210957, -1.380857, -2.552934, -0.778598, 1.570796, 1.781753],accel_mss,speed_ms,0,blend_radius_m)
  movel([0.212521, -1.380569, -2.553139, -0.778681, 1.570796, 1.783318],accel_mss,speed_ms,0,blend_radius_m)
  movel([0.215084, -1.380107, -2.553468, -0.778814, 1.570796, 1.785881],accel_mss,speed_ms,0,blend_radius_m)
  speed_ms = 0.003
  movel([0.215084, -1.367713, -2.547382, -0.797294, 1.570796, 1.785881],accel_mss,speed_ms,0,blend_radius_m)
  speed_ms = 0.01
  movel([0.215084, -1.343947, -2.534831, -0.833611, 1.570796, 1.785881],accel_mss,speed_ms,0,blend_radius_m)
  movel([0.219190, -1.341633, -2.536387, -0.834368, 1.570796, 1.789986],accel_mss,speed_ms,0,blend_radius_m)
  movel([0.219190, -1.365436, -2.548968, -0.797985, 1.570796, 1.789986],accel_mss,speed_ms,0,blend_radius_m)
  speed_ms = 0.003
  movel([0.219190, -1.374715, -2.553555, -0.784120, 1.570796, 1.789986],accel_mss,speed_ms,0,blend_radius_m)
  speed_ms = 0.007
  movel([0.219069, -1.374352, -2.553810, -0.784227, 1.570796, 1.789866],accel_mss,speed_ms,0,blend_radius_m)
  movel([0.218967, -1.373983, -2.554070, -0.784337, 1.570796, 1.789763],accel_mss,speed_ms,0,blend_radius_m)
  movel([0.218876, -1.373591, -2.554345, -0.784453, 1.570796, 1.789672],accel_mss,speed_ms,0,blend_radius_m)
  movel([0.218801, -1.373193, -2.554625, -0.784571, 1.570796, 1.789597],accel_mss,speed_ms,0,blend_radius_m)
  movel([0.218773, -1.372982, -2.554772, -0.784634, 1.570796, 1.789569],accel_mss,speed_ms,0,blend_radius_m)
  movel([0.218757, -1.372770, -2.554922, -0.784698, 1.570796, 1.789553],accel_mss,speed_ms,0,blend_radius_m)
  movel([0.218752, -1.372551, -2.555075, -0.784763, 1.570796, 1.789548],accel_mss,speed_ms,0,blend_radius_m)
  movel([0.218761, -1.372293, -2.555256, -0.784840, 1.570796, 1.789557],accel_mss,speed_ms,0,blend_radius_m)
  movel([0.218780, -1.372029, -2.555441, -0.784919, 1.570796, 1.789577],accel_mss,speed_ms,0,blend_radius_m)
  movel([0.218812, -1.371762, -2.555628, -0.784999, 1.570796, 1.789609],accel_mss,speed_ms,0,blend_radius_m)
  movel([0.218856, -1.371494, -2.555816, -0.785080, 1.570796, 1.789652],accel_mss,speed_ms,0,blend_radius_m)
  movel([0.218910, -1.371221, -2.556006, -0.785162, 1.570796, 1.789707],accel_mss,speed_ms,0,blend_radius_m)
  movel([0.218977, -1.370946, -2.556198, -0.785244, 1.570796, 1.789773],accel_mss,speed_ms,0,blend_radius_m)
  movel([0.219052, -1.370674, -2.556389, -0.785326, 1.570796, 1.789848],accel_mss,speed_ms,0,blend_radius_m)
  movel([0.219139, -1.370400, -2.556580, -0.785409, 1.570796, 1.789936],accel_mss,speed_ms,0,blend_radius_m)
  movel([0.219236, -1.370123, -2.556773, -0.785493, 1.570796, 1.790033],accel_mss,speed_ms,0,blend_radius_m)
  movel([0.219343, -1.369854, -2.556961, -0.785574, 1.570796, 1.790140],accel_mss,speed_ms,0,blend_radius_m)
  movel([0.219460, -1.369584, -2.557149, -0.785656, 1.570796, 1.790256],accel_mss,speed_ms,0,blend_radius_m)
  movel([0.219588, -1.369313, -2.557338, -0.785738, 1.570796, 1.790385],accel_mss,speed_ms,0,blend_radius_m)
  movel([0.219725, -1.369046, -2.557524, -0.785819, 1.570796, 1.790521],accel_mss,speed_ms,0,blend_radius_m)
  movel([0.219873, -1.368780, -2.557710, -0.785900, 1.570796, 1.790670],accel_mss,speed_ms,0,blend_radius_m)
  movel([0.220033, -1.368515, -2.557894, -0.785980, 1.570796, 1.790829],accel_mss,speed_ms,0,blend_radius_m)
  movel([0.220335, -1.368047, -2.558219, -0.786123, 1.570796, 1.791132],accel_mss,speed_ms,0,blend_radius_m)
  movel([0.220651, -1.367583, -2.558541, -0.786265, 1.570796, 1.791447],accel_mss,speed_ms,0,blend_radius_m)
  movel([0.220974, -1.367136, -2.558851, -0.786401, 1.570796, 1.791770],accel_mss,speed_ms,0,blend_radius_m)
  movel([0.221310, -1.366696, -2.559157, -0.786537, 1.570796, 1.792106],accel_mss,speed_ms,0,blend_radius_m)
  movel([0.221486, -1.366479, -2.559307, -0.786603, 1.570796, 1.792283],accel_mss,speed_ms,0,blend_radius_m)
  movel([0.221673, -1.366268, -2.559453, -0.786668, 1.570796, 1.792470],accel_mss,speed_ms,0,blend_radius_m)
  movel([0.221868, -1.366063, -2.559595, -0.786731, 1.570796, 1.792665],accel_mss,speed_ms,0,blend_radius_m)
  movel([0.222292, -1.365637, -2.559890, -0.786862, 1.570796, 1.793089],accel_mss,speed_ms,0,blend_radius_m)
  movel([0.226026, -1.365062, -2.560287, -0.787040, 1.570796, 1.796822],accel_mss,speed_ms,0,blend_radius_m)
  movel([0.229756, -1.364499, -2.560676, -0.787214, 1.570796, 1.800552],accel_mss,speed_ms,0,blend_radius_m)
  movel([0.228572, -1.369199, -2.557418, -0.785773, 1.570796, 1.799368],accel_mss,speed_ms,0,blend_radius_m)
  movel([0.227400, -1.373865, -2.554152, -0.784371, 1.570796, 1.798197],accel_mss,speed_ms,0,blend_radius_m)
  movel([0.223495, -1.374607, -2.553631, -0.784152, 1.570796, 1.794292],accel_mss,speed_ms,0,blend_radius_m)
  movel([0.219589, -1.375360, -2.553100, -0.783929, 1.570796, 1.790385],accel_mss,speed_ms,0,blend_radius_m)
  movel([0.219418, -1.375139, -2.553256, -0.783994, 1.570796, 1.790214],accel_mss,speed_ms,0,blend_radius_m)
  movel([0.219327, -1.375008, -2.553348, -0.784033, 1.570796, 1.790123],accel_mss,speed_ms,0,blend_radius_m)
  movel([0.219251, -1.374866, -2.553448, -0.784075, 1.570796, 1.790047],accel_mss,speed_ms,0,blend_radius_m)
  movel([0.219190, -1.374715, -2.553555, -0.784120, 1.570796, 1.789986],accel_mss,speed_ms,0,blend_radius_m)
  speed_ms = 0.003
  movel([0.219190, -1.377851, -2.555068, -0.779471, 1.570796, 1.789986],accel_mss,speed_ms,0,blend_radius_m)
  speed_ms = 0.007
  movel([0.219069, -1.377489, -2.555323, -0.779577, 1.570796, 1.789866],accel_mss,speed_ms,0,blend_radius_m)
  movel([0.218967, -1.377120, -2.555584, -0.779685, 1.570796, 1.789763],accel_mss,speed_ms,0,blend_radius_m)
  movel([0.218876, -1.376730, -2.555859, -0.779799, 1.570796, 1.789672],accel_mss,speed_ms,0,blend_radius_m)
  movel([0.218801, -1.376333, -2.556140, -0.779916, 1.570796, 1.789597],accel_mss,speed_ms,0,blend_radius_m)
  movel([0.218773, -1.376123, -2.556288, -0.779978, 1.570796, 1.789569],accel_mss,speed_ms,0,blend_radius_m)
  movel([0.218757, -1.375910, -2.556438, -0.780041, 1.570796, 1.789553],accel_mss,speed_ms,0,blend_radius_m)
  movel([0.218752, -1.375692, -2.556592, -0.780105, 1.570796, 1.789548],accel_mss,speed_ms,0,blend_radius_m)
  movel([0.218761, -1.375435, -2.556773, -0.780182, 1.570796, 1.789557],accel_mss,speed_ms,0,blend_radius_m)
  movel([0.218780, -1.375171, -2.556958, -0.780260, 1.570796, 1.789577],accel_mss,speed_ms,0,blend_radius_m)
  movel([0.218812, -1.374906, -2.557145, -0.780338, 1.570796, 1.789609],accel_mss,speed_ms,0,blend_radius_m)
  movel([0.218856, -1.374638, -2.557334, -0.780418, 1.570796, 1.789652],accel_mss,speed_ms,0,blend_radius_m)
  movel([0.218910, -1.374366, -2.557525, -0.780499, 1.570796, 1.789707],accel_mss,speed_ms,0,blend_radius_m)
  movel([0.218977, -1.374091, -2.557717, -0.780580, 1.570796, 1.789773],accel_mss,speed_ms,0,blend_radius_m)
  movel([0.219052, -1.373820, -2.557908, -0.780661, 1.570796, 1.789848],accel_mss,speed_ms,0,blend_radius_m)
  movel([0.219139, -1.373546, -2.558100, -0.780743, 1.570796, 1.789936],accel_mss,speed_ms,0,blend_radius_m)
  movel([0.219236, -1.373270, -2.558293, -0.780825, 1.570796, 1.790033],accel_mss,speed_ms,0,blend_radius_m)
  movel([0.219343, -1.373001, -2.558482, -0.780906, 1.570796, 1.790140],accel_mss,speed_ms,0,blend_radius_m)
  movel([0.219460, -1.372733, -2.558670, -0.780986, 1.570796, 1.790256],accel_mss,speed_ms,0,blend_radius_m)
  movel([0.219588, -1.372462, -2.558860, -0.781067, 1.570796, 1.790385],accel_mss,speed_ms,0,blend_radius_m)
  movel([0.219725, -1.372196, -2.559046, -0.781147, 1.570796, 1.790521],accel_mss,speed_ms,0,blend_radius_m)
  movel([0.219873, -1.371930, -2.559232, -0.781227, 1.570796, 1.790670],accel_mss,speed_ms,0,blend_radius_m)
  movel([0.220033, -1.371666, -2.559416, -0.781307, 1.570796, 1.790829],accel_mss,speed_ms,0,blend_radius_m)
  movel([0.220335, -1.371199, -2.559743, -0.781448, 1.570796, 1.791132],accel_mss,speed_ms,0,blend_radius_m)
  movel([0.220651, -1.370736, -2.560066, -0.781587, 1.570796, 1.791447],accel_mss,speed_ms,0,blend_radius_m)
  movel([0.220974, -1.370290, -2.560376, -0.781722, 1.570796, 1.791770],accel_mss,speed_ms,0,blend_radius_m)
  movel([0.221310, -1.369851, -2.560682, -0.781856, 1.570796, 1.792106],accel_mss,speed_ms,0,blend_radius_m)
  movel([0.221486, -1.369635, -2.560833, -0.781921, 1.570796, 1.792283],accel_mss,speed_ms,0,blend_radius_m)
  movel([0.221673, -1.369424, -2.560980, -0.781986, 1.570796, 1.792470],accel_mss,speed_ms,0,blend_radius_m)
  movel([0.221868, -1.369220, -2.561122, -0.782048, 1.570796, 1.792665],accel_mss,speed_ms,0,blend_radius_m)
  movel([0.222292, -1.368794, -2.561417, -0.782177, 1.570796, 1.793089],accel_mss,speed_ms,0,blend_radius_m)
  movel([0.226026, -1.368221, -2.561816, -0.782353, 1.570796, 1.796822],accel_mss,speed_ms,0,blend_radius_m)
  movel([0.229756, -1.367659, -2.562205, -0.782525, 1.570796, 1.800552],accel_mss,speed_ms,0,blend_radius_m)
  movel([0.228572, -1.372348, -2.558940, -0.781102, 1.570796, 1.799368],accel_mss,speed_ms,0,blend_radius_m)
  movel([0.227400, -1.377003, -2.555666, -0.779719, 1.570796, 1.798197],accel_mss,speed_ms,0,blend_radius_m)
  movel([0.223495, -1.377743, -2.555144, -0.779502, 1.570796, 1.794292],accel_mss,speed_ms,0,blend_radius_m)
  movel([0.219589, -1.378494, -2.554612, -0.779283, 1.570796, 1.790385],accel_mss,speed_ms,0,blend_radius_m)
  movel([0.219418, -1.378274, -2.554768, -0.779347, 1.570796, 1.790214],accel_mss,speed_ms,0,blend_radius_m)
  movel([0.219327, -1.378143, -2.554861, -0.779385, 1.570796, 1.790123],accel_mss,speed_ms,0,blend_radius_m)
  movel([0.219251, -1.378001, -2.554961, -0.779427, 1.570796, 1.790047],accel_mss,speed_ms,0,blend_radius_m)
  movel([0.219190, -1.377851, -2.555068, -0.779471, 1.570796, 1.789986],accel_mss,speed_ms,0,blend_radius_m)
  speed_ms = 0.003
  movel([0.219190, -1.365436, -2.548968, -0.797985, 1.570796, 1.789986],accel_mss,speed_ms,0,blend_radius_m)
  speed_ms = 0.01
  movel([0.219190, -1.341633, -2.536387, -0.834368, 1.570796, 1.789986],accel_mss,speed_ms,0,blend_radius_m)
  movel([0.211822, -1.348948, -2.531442, -0.831999, 1.570796, 1.782619],accel_mss,speed_ms,0,blend_radius_m)
  movel([0.211822, -1.372635, -2.543931, -0.795823, 1.570796, 1.782619],accel_mss,speed_ms,0,blend_radius_m)
  speed_ms = 0.003
  movel([0.211822, -1.381864, -2.548484, -0.782041, 1.570796, 1.782619],accel_mss,speed_ms,0,blend_radius_m)
  speed_ms = 0.007
  movel([0.210818, -1.385912, -2.545582, -0.780896, 1.570796, 1.781615],accel_mss,speed_ms,0,blend_radius_m)
  movel([0.210430, -1.387463, -2.544463, -0.780463, 1.570796, 1.781227],accel_mss,speed_ms,0,blend_radius_m)
  movel([0.210091, -1.388779, -2.543511, -0.780099, 1.570796, 1.780887],accel_mss,speed_ms,0,blend_radius_m)
  movel([0.209783, -1.389944, -2.542667, -0.779778, 1.570796, 1.780579],accel_mss,speed_ms,0,blend_radius_m)
  movel([0.209765, -1.389982, -2.542639, -0.779768, 1.570796, 1.780561],accel_mss,speed_ms,0,blend_radius_m)
  movel([0.209734, -1.390017, -2.542614, -0.779758, 1.570796, 1.780530],accel_mss,speed_ms,0,blend_radius_m)
  movel([0.209698, -1.390044, -2.542594, -0.779751, 1.570796, 1.780494],accel_mss,speed_ms,0,blend_radius_m)
  movel([0.209659, -1.390066, -2.542579, -0.779745, 1.570796, 1.780455],accel_mss,speed_ms,0,blend_radius_m)
  movel([0.209103, -1.390320, -2.542394, -0.779675, 1.570796, 1.779899],accel_mss,speed_ms,0,blend_radius_m)
  movel([0.208458, -1.390611, -2.542183, -0.779596, 1.570796, 1.779255],accel_mss,speed_ms,0,blend_radius_m)
  movel([0.207710, -1.390939, -2.541944, -0.779506, 1.570796, 1.778507],accel_mss,speed_ms,0,blend_radius_m)
  movel([0.205779, -1.391779, -2.541333, -0.779277, 1.570796, 1.776575],accel_mss,speed_ms,0,blend_radius_m)
  movel([0.205514, -1.392938, -2.540488, -0.778963, 1.570796, 1.776310],accel_mss,speed_ms,0,blend_radius_m)
  movel([0.205249, -1.394094, -2.539643, -0.778652, 1.570796, 1.776046],accel_mss,speed_ms,0,blend_radius_m)
  movel([0.203680, -1.394883, -2.539065, -0.778441, 1.570796, 1.774476],accel_mss,speed_ms,0,blend_radius_m)
  movel([0.202110, -1.395671, -2.538487, -0.778231, 1.570796, 1.772906],accel_mss,speed_ms,0,blend_radius_m)
  movel([0.201949, -1.396236, -2.538072, -0.778080, 1.570796, 1.772745],accel_mss,speed_ms,0,blend_radius_m)
  movel([0.201788, -1.396801, -2.537657, -0.777931, 1.570796, 1.772584],accel_mss,speed_ms,0,blend_radius_m)
  movel([0.186663, -1.399616, -2.535581, -0.777192, 1.570796, 1.757460],accel_mss,speed_ms,0,blend_radius_m)
  movel([0.171550, -1.402607, -2.533363, -0.776419, 1.570796, 1.742347],accel_mss,speed_ms,0,blend_radius_m)
  movel([0.171931, -1.402198, -2.533667, -0.776524, 1.570796, 1.742727],accel_mss,speed_ms,0,blend_radius_m)
  movel([0.172504, -1.401569, -2.534134, -0.776686, 1.570796, 1.743301],accel_mss,speed_ms,0,blend_radius_m)
  movel([0.173060, -1.400927, -2.534611, -0.776852, 1.570796, 1.743857],accel_mss,speed_ms,0,blend_radius_m)
  movel([0.173596, -1.400274, -2.535094, -0.777021, 1.570796, 1.744393],accel_mss,speed_ms,0,blend_radius_m)
  movel([0.174083, -1.399647, -2.535558, -0.777184, 1.570796, 1.744879],accel_mss,speed_ms,0,blend_radius_m)
  movel([0.174543, -1.399012, -2.536027, -0.777349, 1.570796, 1.745340],accel_mss,speed_ms,0,blend_radius_m)
  movel([0.174979, -1.398368, -2.536503, -0.777518, 1.570796, 1.745776],accel_mss,speed_ms,0,blend_radius_m)
  movel([0.175377, -1.397737, -2.536968, -0.777684, 1.570796, 1.746173],accel_mss,speed_ms,0,blend_radius_m)
  movel([0.175746, -1.397099, -2.537438, -0.777852, 1.570796, 1.746543],accel_mss,speed_ms,0,blend_radius_m)
  movel([0.176087, -1.396459, -2.537909, -0.778021, 1.570796, 1.746883],accel_mss,speed_ms,0,blend_radius_m)
  movel([0.176402, -1.395815, -2.538382, -0.778192, 1.570796, 1.747198],accel_mss,speed_ms,0,blend_radius_m)
  movel([0.176687, -1.395168, -2.538857, -0.778365, 1.570796, 1.747484],accel_mss,speed_ms,0,blend_radius_m)
  movel([0.176944, -1.394520, -2.539331, -0.778538, 1.570796, 1.747740],accel_mss,speed_ms,0,blend_radius_m)
  movel([0.177132, -1.393965, -2.539737, -0.778687, 1.570796, 1.747928],accel_mss,speed_ms,0,blend_radius_m)
  movel([0.177282, -1.393416, -2.540138, -0.778834, 1.570796, 1.748078],accel_mss,speed_ms,0,blend_radius_m)
  movel([0.177437, -1.392717, -2.540649, -0.779023, 1.570796, 1.748233],accel_mss,speed_ms,0,blend_radius_m)
  movel([0.177569, -1.392021, -2.541157, -0.779212, 1.570796, 1.748365],accel_mss,speed_ms,0,blend_radius_m)
  movel([0.177678, -1.391326, -2.541663, -0.779400, 1.570796, 1.748474],accel_mss,speed_ms,0,blend_radius_m)
  movel([0.177765, -1.390635, -2.542165, -0.779589, 1.570796, 1.748561],accel_mss,speed_ms,0,blend_radius_m)
  movel([0.177804, -1.390095, -2.542557, -0.779737, 1.570796, 1.748600],accel_mss,speed_ms,0,blend_radius_m)
  movel([0.177803, -1.389568, -2.542940, -0.779881, 1.570796, 1.748600],accel_mss,speed_ms,0,blend_radius_m)
  movel([0.177770, -1.389022, -2.543335, -0.780032, 1.570796, 1.748566],accel_mss,speed_ms,0,blend_radius_m)
  movel([0.177709, -1.388485, -2.543724, -0.780180, 1.570796, 1.748505],accel_mss,speed_ms,0,blend_radius_m)
  movel([0.177623, -1.387960, -2.544104, -0.780325, 1.570796, 1.748419],accel_mss,speed_ms,0,blend_radius_m)
  movel([0.177507, -1.387444, -2.544477, -0.780468, 1.570796, 1.748303],accel_mss,speed_ms,0,blend_radius_m)
  movel([0.177367, -1.386941, -2.544839, -0.780608, 1.570796, 1.748164],accel_mss,speed_ms,0,blend_radius_m)
  movel([0.177202, -1.386452, -2.545192, -0.780745, 1.570796, 1.747998],accel_mss,speed_ms,0,blend_radius_m)
  movel([0.177016, -1.385996, -2.545521, -0.780872, 1.570796, 1.747812],accel_mss,speed_ms,0,blend_radius_m)
  movel([0.176805, -1.385557, -2.545837, -0.780995, 1.570796, 1.747602],accel_mss,speed_ms,0,blend_radius_m)
  movel([0.176571, -1.385133, -2.546142, -0.781114, 1.570796, 1.747367],accel_mss,speed_ms,0,blend_radius_m)
  movel([0.176332, -1.384764, -2.546407, -0.781218, 1.570796, 1.747129],accel_mss,speed_ms,0,blend_radius_m)
  movel([0.176063, -1.384418, -2.546656, -0.781316, 1.570796, 1.746860],accel_mss,speed_ms,0,blend_radius_m)
  movel([0.175766, -1.384096, -2.546886, -0.781406, 1.570796, 1.746563],accel_mss,speed_ms,0,blend_radius_m)
  movel([0.175624, -1.383951, -2.546991, -0.781447, 1.570796, 1.746420],accel_mss,speed_ms,0,blend_radius_m)
  movel([0.175484, -1.383805, -2.547095, -0.781489, 1.570796, 1.746280],accel_mss,speed_ms,0,blend_radius_m)
  movel([0.175366, -1.383675, -2.547188, -0.781525, 1.570796, 1.746162],accel_mss,speed_ms,0,blend_radius_m)
  movel([0.175294, -1.383592, -2.547248, -0.781549, 1.570796, 1.746091],accel_mss,speed_ms,0,blend_radius_m)
  movel([0.175286, -1.383565, -2.547267, -0.781557, 1.570796, 1.746082],accel_mss,speed_ms,0,blend_radius_m)
  movel([0.175293, -1.383530, -2.547292, -0.781567, 1.570796, 1.746089],accel_mss,speed_ms,0,blend_radius_m)
  movel([0.175316, -1.383496, -2.547317, -0.781576, 1.570796, 1.746112],accel_mss,speed_ms,0,blend_radius_m)
  movel([0.175349, -1.383468, -2.547337, -0.781584, 1.570796, 1.746145],accel_mss,speed_ms,0,blend_radius_m)
  movel([0.175387, -1.383452, -2.547348, -0.781589, 1.570796, 1.746183],accel_mss,speed_ms,0,blend_radius_m)
  movel([0.176404, -1.383221, -2.547514, -0.781654, 1.570796, 1.747200],accel_mss,speed_ms,0,blend_radius_m)
  movel([0.177420, -1.382995, -2.547675, -0.781718, 1.570796, 1.748216],accel_mss,speed_ms,0,blend_radius_m)
  movel([0.179187, -1.382613, -2.547949, -0.781827, 1.570796, 1.749983],accel_mss,speed_ms,0,blend_radius_m)
  movel([0.180950, -1.382244, -2.548213, -0.781932, 1.570796, 1.751746],accel_mss,speed_ms,0,blend_radius_m)
  movel([0.190746, -1.380271, -2.549621, -0.782498, 1.570796, 1.761543],accel_mss,speed_ms,0,blend_radius_m)
  movel([0.206333, -1.377291, -2.551736, -0.783362, 1.570796, 1.777129],accel_mss,speed_ms,0,blend_radius_m)
  movel([0.206200, -1.378024, -2.551216, -0.783148, 1.570796, 1.776996],accel_mss,speed_ms,0,blend_radius_m)
  movel([0.206065, -1.378755, -2.550698, -0.782936, 1.570796, 1.776862],accel_mss,speed_ms,0,blend_radius_m)
  movel([0.207335, -1.379009, -2.550518, -0.782862, 1.570796, 1.778131],accel_mss,speed_ms,0,blend_radius_m)
  movel([0.208603, -1.379265, -2.550336, -0.782788, 1.570796, 1.779399],accel_mss,speed_ms,0,blend_radius_m)
  movel([0.208397, -1.380302, -2.549598, -0.782489, 1.570796, 1.779194],accel_mss,speed_ms,0,blend_radius_m)
  movel([0.208190, -1.381339, -2.548859, -0.782191, 1.570796, 1.778987],accel_mss,speed_ms,0,blend_radius_m)
  movel([0.209668, -1.381528, -2.548724, -0.782137, 1.570796, 1.780464],accel_mss,speed_ms,0,blend_radius_m)
  movel([0.210257, -1.381605, -2.548669, -0.782115, 1.570796, 1.781053],accel_mss,speed_ms,0,blend_radius_m)
  movel([0.210809, -1.381683, -2.548613, -0.782092, 1.570796, 1.781606],accel_mss,speed_ms,0,blend_radius_m)
  movel([0.211272, -1.381752, -2.548564, -0.782073, 1.570796, 1.782068],accel_mss,speed_ms,0,blend_radius_m)
  movel([0.211483, -1.381790, -2.548537, -0.782062, 1.570796, 1.782280],accel_mss,speed_ms,0,blend_radius_m)
  movel([0.211822, -1.381864, -2.548484, -0.782041, 1.570796, 1.782619],accel_mss,speed_ms,0,blend_radius_m)
  speed_ms = 0.003
  movel([0.211822, -1.384983, -2.549985, -0.777420, 1.570796, 1.782619],accel_mss,speed_ms,0,blend_radius_m)
  speed_ms = 0.007
  movel([0.210818, -1.389020, -2.547077, -0.776292, 1.570796, 1.781615],accel_mss,speed_ms,0,blend_radius_m)
  movel([0.210430, -1.390568, -2.545956, -0.775866, 1.570796, 1.781227],accel_mss,speed_ms,0,blend_radius_m)
  movel([0.210091, -1.391881, -2.545002, -0.775506, 1.570796, 1.780887],accel_mss,speed_ms,0,blend_radius_m)
  movel([0.209783, -1.393043, -2.544156, -0.775191, 1.570796, 1.780579],accel_mss,speed_ms,0,blend_radius_m)
  movel([0.209765, -1.393081, -2.544128, -0.775180, 1.570796, 1.780561],accel_mss,speed_ms,0,blend_radius_m)
  movel([0.209734, -1.393116, -2.544102, -0.775171, 1.570796, 1.780530],accel_mss,speed_ms,0,blend_radius_m)
  movel([0.209698, -1.393143, -2.544083, -0.775164, 1.570796, 1.780494],accel_mss,speed_ms,0,blend_radius_m)
  movel([0.209659, -1.393164, -2.544067, -0.775158, 1.570796, 1.780455],accel_mss,speed_ms,0,blend_radius_m)
  movel([0.209103, -1.393418, -2.543882, -0.775089, 1.570796, 1.779899],accel_mss,speed_ms,0,blend_radius_m)
  movel([0.208458, -1.393708, -2.543670, -0.775011, 1.570796, 1.779255],accel_mss,speed_ms,0,blend_radius_m)
  movel([0.207710, -1.394035, -2.543431, -0.774923, 1.570796, 1.778507],accel_mss,speed_ms,0,blend_radius_m)
  movel([0.205779, -1.394873, -2.542818, -0.774697, 1.570796, 1.776575],accel_mss,speed_ms,0,blend_radius_m)
  movel([0.205514, -1.396029, -2.541972, -0.774388, 1.570796, 1.776310],accel_mss,speed_ms,0,blend_radius_m)
  movel([0.205249, -1.397183, -2.541125, -0.774081, 1.570796, 1.776046],accel_mss,speed_ms,0,blend_radius_m)
  movel([0.203680, -1.397970, -2.540546, -0.773873, 1.570796, 1.774476],accel_mss,speed_ms,0,blend_radius_m)
  movel([0.202110, -1.398756, -2.539967, -0.773666, 1.570796, 1.772906],accel_mss,speed_ms,0,blend_radius_m)
  movel([0.201949, -1.399319, -2.539551, -0.773519, 1.570796, 1.772745],accel_mss,speed_ms,0,blend_radius_m)
  movel([0.201788, -1.399883, -2.539135, -0.773371, 1.570796, 1.772584],accel_mss,speed_ms,0,blend_radius_m)
  movel([0.186663, -1.402690, -2.537054, -0.772644, 1.570796, 1.757460],accel_mss,speed_ms,0,blend_radius_m)
  movel([0.171550, -1.405674, -2.534831, -0.771884, 1.570796, 1.742347],accel_mss,speed_ms,0,blend_radius_m)
  movel([0.171931, -1.405266, -2.535136, -0.771987, 1.570796, 1.742727],accel_mss,speed_ms,0,blend_radius_m)
  movel([0.172504, -1.404639, -2.535604, -0.772146, 1.570796, 1.743301],accel_mss,speed_ms,0,blend_radius_m)
  movel([0.173060, -1.403998, -2.536082, -0.772309, 1.570796, 1.743857],accel_mss,speed_ms,0,blend_radius_m)
  movel([0.173596, -1.403347, -2.536567, -0.772476, 1.570796, 1.744393],accel_mss,speed_ms,0,blend_radius_m)
  movel([0.174083, -1.402721, -2.537032, -0.772636, 1.570796, 1.744879],accel_mss,speed_ms,0,blend_radius_m)
  movel([0.174543, -1.402088, -2.537502, -0.772799, 1.570796, 1.745340],accel_mss,speed_ms,0,blend_radius_m)
  movel([0.174979, -1.401446, -2.537978, -0.772965, 1.570796, 1.745776],accel_mss,speed_ms,0,blend_radius_m)
  movel([0.175377, -1.400817, -2.538444, -0.773128, 1.570796, 1.746173],accel_mss,speed_ms,0,blend_radius_m)
  movel([0.175746, -1.400180, -2.538915, -0.773294, 1.570796, 1.746543],accel_mss,speed_ms,0,blend_radius_m)
  movel([0.176087, -1.399541, -2.539387, -0.773461, 1.570796, 1.746883],accel_mss,speed_ms,0,blend_radius_m)
  movel([0.176402, -1.398899, -2.539861, -0.773629, 1.570796, 1.747198],accel_mss,speed_ms,0,blend_radius_m)
  movel([0.176687, -1.398253, -2.540337, -0.773799, 1.570796, 1.747484],accel_mss,speed_ms,0,blend_radius_m)
  movel([0.176944, -1.397607, -2.540813, -0.773969, 1.570796, 1.747740],accel_mss,speed_ms,0,blend_radius_m)
  movel([0.177132, -1.397054, -2.541219, -0.774116, 1.570796, 1.747928],accel_mss,speed_ms,0,blend_radius_m)
  movel([0.177282, -1.396506, -2.541622, -0.774261, 1.570796, 1.748078],accel_mss,speed_ms,0,blend_radius_m)
  movel([0.177437, -1.395809, -2.542133, -0.774447, 1.570796, 1.748233],accel_mss,speed_ms,0,blend_radius_m)
  movel([0.177569, -1.395114, -2.542642, -0.774633, 1.570796, 1.748365],accel_mss,speed_ms,0,blend_radius_m)
  movel([0.177678, -1.394421, -2.543149, -0.774819, 1.570796, 1.748474],accel_mss,speed_ms,0,blend_radius_m)
  movel([0.177765, -1.393732, -2.543653, -0.775004, 1.570796, 1.748561],accel_mss,speed_ms,0,blend_radius_m)
  movel([0.177804, -1.393194, -2.544045, -0.775150, 1.570796, 1.748600],accel_mss,speed_ms,0,blend_radius_m)
  movel([0.177803, -1.392668, -2.544429, -0.775292, 1.570796, 1.748600],accel_mss,speed_ms,0,blend_radius_m)
  movel([0.177770, -1.392123, -2.544826, -0.775440, 1.570796, 1.748566],accel_mss,speed_ms,0,blend_radius_m)
  movel([0.177709, -1.391588, -2.545215, -0.775586, 1.570796, 1.748505],accel_mss,speed_ms,0,blend_radius_m)
  movel([0.177623, -1.391064, -2.545596, -0.775730, 1.570796, 1.748419],accel_mss,speed_ms,0,blend_radius_m)
  movel([0.177507, -1.390549, -2.545969, -0.775871, 1.570796, 1.748303],accel_mss,speed_ms,0,blend_radius_m)
  movel([0.177367, -1.390048, -2.546333, -0.776008, 1.570796, 1.748164],accel_mss,speed_ms,0,blend_radius_m)
  movel([0.177202, -1.389559, -2.546687, -0.776143, 1.570796, 1.747998],accel_mss,speed_ms,0,blend_radius_m)
  movel([0.177016, -1.389104, -2.547016, -0.776269, 1.570796, 1.747812],accel_mss,speed_ms,0,blend_radius_m)
  movel([0.176805, -1.388666, -2.547333, -0.776390, 1.570796, 1.747602],accel_mss,speed_ms,0,blend_radius_m)
  movel([0.176571, -1.388243, -2.547638, -0.776507, 1.570796, 1.747367],accel_mss,speed_ms,0,blend_radius_m)
  movel([0.176332, -1.387875, -2.547904, -0.776610, 1.570796, 1.747129],accel_mss,speed_ms,0,blend_radius_m)
  movel([0.176063, -1.387530, -2.548153, -0.776706, 1.570796, 1.746860],accel_mss,speed_ms,0,blend_radius_m)
  movel([0.175766, -1.387209, -2.548384, -0.776795, 1.570796, 1.746563],accel_mss,speed_ms,0,blend_radius_m)
  movel([0.175624, -1.387064, -2.548489, -0.776836, 1.570796, 1.746420],accel_mss,speed_ms,0,blend_radius_m)
  movel([0.175484, -1.386919, -2.548594, -0.776876, 1.570796, 1.746280],accel_mss,speed_ms,0,blend_radius_m)
  movel([0.175366, -1.386790, -2.548687, -0.776913, 1.570796, 1.746162],accel_mss,speed_ms,0,blend_radius_m)
  movel([0.175294, -1.386707, -2.548746, -0.776936, 1.570796, 1.746091],accel_mss,speed_ms,0,blend_radius_m)
  movel([0.175286, -1.386679, -2.548766, -0.776943, 1.570796, 1.746082],accel_mss,speed_ms,0,blend_radius_m)
  movel([0.175293, -1.386645, -2.548791, -0.776953, 1.570796, 1.746089],accel_mss,speed_ms,0,blend_radius_m)
  movel([0.175316, -1.386611, -2.548815, -0.776963, 1.570796, 1.746112],accel_mss,speed_ms,0,blend_radius_m)
  movel([0.175349, -1.386583, -2.548835, -0.776970, 1.570796, 1.746145],accel_mss,speed_ms,0,blend_radius_m)
  movel([0.175387, -1.386567, -2.548847, -0.776975, 1.570796, 1.746183],accel_mss,speed_ms,0,blend_radius_m)
  movel([0.176404, -1.386336, -2.549013, -0.777040, 1.570796, 1.747200],accel_mss,speed_ms,0,blend_radius_m)
  movel([0.177420, -1.386111, -2.549175, -0.777103, 1.570796, 1.748216],accel_mss,speed_ms,0,blend_radius_m)
  movel([0.179187, -1.385730, -2.549449, -0.777210, 1.570796, 1.749983],accel_mss,speed_ms,0,blend_radius_m)
  movel([0.180950, -1.385362, -2.549713, -0.777314, 1.570796, 1.751746],accel_mss,speed_ms,0,blend_radius_m)
  movel([0.190746, -1.383393, -2.551125, -0.777871, 1.570796, 1.761543],accel_mss,speed_ms,0,blend_radius_m)
  movel([0.206333, -1.380421, -2.553244, -0.778724, 1.570796, 1.777129],accel_mss,speed_ms,0,blend_radius_m)
  movel([0.206200, -1.381152, -2.552724, -0.778513, 1.570796, 1.776996],accel_mss,speed_ms,0,blend_radius_m)
  movel([0.206065, -1.381881, -2.552205, -0.778303, 1.570796, 1.776862],accel_mss,speed_ms,0,blend_radius_m)
  movel([0.207335, -1.382135, -2.552024, -0.778231, 1.570796, 1.778131],accel_mss,speed_ms,0,blend_radius_m)
  movel([0.208603, -1.382390, -2.551841, -0.778158, 1.570796, 1.779399],accel_mss,speed_ms,0,blend_radius_m)
  movel([0.208397, -1.383425, -2.551102, -0.777862, 1.570796, 1.779194],accel_mss,speed_ms,0,blend_radius_m)
  movel([0.208190, -1.384459, -2.550362, -0.777569, 1.570796, 1.778987],accel_mss,speed_ms,0,blend_radius_m)
  movel([0.209668, -1.384648, -2.550226, -0.777515, 1.570796, 1.780464],accel_mss,speed_ms,0,blend_radius_m)
  movel([0.210257, -1.384725, -2.550171, -0.777493, 1.570796, 1.781053],accel_mss,speed_ms,0,blend_radius_m)
  movel([0.210809, -1.384802, -2.550115, -0.777472, 1.570796, 1.781606],accel_mss,speed_ms,0,blend_radius_m)
  movel([0.211272, -1.384871, -2.550066, -0.777452, 1.570796, 1.782068],accel_mss,speed_ms,0,blend_radius_m)
  movel([0.211483, -1.384909, -2.550039, -0.777441, 1.570796, 1.782280],accel_mss,speed_ms,0,blend_radius_m)
  movel([0.211822, -1.384983, -2.549985, -0.777420, 1.570796, 1.782619],accel_mss,speed_ms,0,blend_radius_m)
  speed_ms = 0.003
  movel([0.211822, -1.372635, -2.543931, -0.795823, 1.570796, 1.782619],accel_mss,speed_ms,0,blend_radius_m)
  speed_ms = 0.01
  movel([0.211822, -1.348948, -2.531442, -0.831999, 1.570796, 1.782619],accel_mss,speed_ms,0,blend_radius_m)
  movel([0.208233, -1.333772, -2.541623, -0.836993, 1.570796, 1.779029],accel_mss,speed_ms,0,blend_radius_m)
  movel([0.208233, -1.357697, -2.554302, -0.800390, 1.570796, 1.779029],accel_mss,speed_ms,0,blend_radius_m)
  speed_ms = 0.003
  movel([0.208233, -1.367028, -2.558926, -0.786435, 1.570796, 1.779029],accel_mss,speed_ms,0,blend_radius_m)
  speed_ms = 0.007
  movel([0.192461, -1.370092, -2.556795, -0.785502, 1.570796, 1.763257],accel_mss,speed_ms,0,blend_radius_m)
  movel([0.176700, -1.373348, -2.554516, -0.784525, 1.570796, 1.747496],accel_mss,speed_ms,0,blend_radius_m)
  movel([0.177720, -1.372310, -2.555244, -0.784835, 1.570796, 1.748516],accel_mss,speed_ms,0,blend_radius_m)
  movel([0.178177, -1.371836, -2.555576, -0.784977, 1.570796, 1.748973],accel_mss,speed_ms,0,blend_radius_m)
  movel([0.178623, -1.371349, -2.555917, -0.785123, 1.570796, 1.749419],accel_mss,speed_ms,0,blend_radius_m)
  movel([0.179054, -1.370857, -2.556261, -0.785271, 1.570796, 1.749850],accel_mss,speed_ms,0,blend_radius_m)
  movel([0.179470, -1.370354, -2.556612, -0.785423, 1.570796, 1.750267],accel_mss,speed_ms,0,blend_radius_m)
  movel([0.179870, -1.369847, -2.556966, -0.785576, 1.570796, 1.750666],accel_mss,speed_ms,0,blend_radius_m)
  movel([0.180257, -1.369331, -2.557325, -0.785732, 1.570796, 1.751054],accel_mss,speed_ms,0,blend_radius_m)
  movel([0.180628, -1.368810, -2.557688, -0.785891, 1.570796, 1.751424],accel_mss,speed_ms,0,blend_radius_m)
  movel([0.180979, -1.368291, -2.558050, -0.786049, 1.570796, 1.751775],accel_mss,speed_ms,0,blend_radius_m)
  movel([0.181310, -1.367767, -2.558414, -0.786209, 1.570796, 1.752107],accel_mss,speed_ms,0,blend_radius_m)
  movel([0.181624, -1.367240, -2.558780, -0.786370, 1.570796, 1.752420],accel_mss,speed_ms,0,blend_radius_m)
  movel([0.181922, -1.366707, -2.559149, -0.786533, 1.570796, 1.752718],accel_mss,speed_ms,0,blend_radius_m)
  movel([0.182200, -1.366174, -2.559518, -0.786697, 1.570796, 1.752996],accel_mss,speed_ms,0,blend_radius_m)
  movel([0.182457, -1.365638, -2.559889, -0.786862, 1.570796, 1.753253],accel_mss,speed_ms,0,blend_radius_m)
  movel([0.182698, -1.365102, -2.560260, -0.787028, 1.570796, 1.753494],accel_mss,speed_ms,0,blend_radius_m)
  movel([0.182918, -1.364562, -2.560632, -0.787195, 1.570796, 1.753714],accel_mss,speed_ms,0,blend_radius_m)
  movel([0.183120, -1.364022, -2.561004, -0.787362, 1.570796, 1.753916],accel_mss,speed_ms,0,blend_radius_m)
  movel([0.183301, -1.363482, -2.561377, -0.787530, 1.570796, 1.754097],accel_mss,speed_ms,0,blend_radius_m)
  movel([0.183460, -1.362946, -2.561745, -0.787697, 1.570796, 1.754256],accel_mss,speed_ms,0,blend_radius_m)
  movel([0.183600, -1.362412, -2.562113, -0.787864, 1.570796, 1.754396],accel_mss,speed_ms,0,blend_radius_m)
  movel([0.183717, -1.361881, -2.562477, -0.788031, 1.570796, 1.754514],accel_mss,speed_ms,0,blend_radius_m)
  movel([0.183813, -1.361356, -2.562838, -0.788196, 1.570796, 1.754609],accel_mss,speed_ms,0,blend_radius_m)
  movel([0.183892, -1.360820, -2.563205, -0.788364, 1.570796, 1.754688],accel_mss,speed_ms,0,blend_radius_m)
  movel([0.183948, -1.360291, -2.563567, -0.788531, 1.570796, 1.754744],accel_mss,speed_ms,0,blend_radius_m)
  movel([0.183986, -1.359767, -2.563925, -0.788697, 1.570796, 1.754782],accel_mss,speed_ms,0,blend_radius_m)
  movel([0.184002, -1.359250, -2.564278, -0.788861, 1.570796, 1.754798],accel_mss,speed_ms,0,blend_radius_m)
  movel([0.183994, -1.358743, -2.564624, -0.789022, 1.570796, 1.754790],accel_mss,speed_ms,0,blend_radius_m)
  movel([0.183968, -1.358240, -2.564967, -0.789182, 1.570796, 1.754765],accel_mss,speed_ms,0,blend_radius_m)
  movel([0.183922, -1.357746, -2.565303, -0.789339, 1.570796, 1.754718],accel_mss,speed_ms,0,blend_radius_m)
  movel([0.183841, -1.357236, -2.565651, -0.789503, 1.570796, 1.754637],accel_mss,speed_ms,0,blend_radius_m)
  movel([0.183722, -1.356746, -2.565984, -0.789660, 1.570796, 1.754519],accel_mss,speed_ms,0,blend_radius_m)
  movel([0.183540, -1.356161, -2.566381, -0.789848, 1.570796, 1.754336],accel_mss,speed_ms,0,blend_radius_m)
  movel([0.183332, -1.355590, -2.566768, -0.790031, 1.570796, 1.754129],accel_mss,speed_ms,0,blend_radius_m)
  movel([0.183103, -1.355040, -2.567140, -0.790209, 1.570796, 1.753900],accel_mss,speed_ms,0,blend_radius_m)
  movel([0.182850, -1.354506, -2.567501, -0.790381, 1.570796, 1.753646],accel_mss,speed_ms,0,blend_radius_m)
  movel([0.182624, -1.354112, -2.567768, -0.790509, 1.570796, 1.753421],accel_mss,speed_ms,0,blend_radius_m)
  movel([0.182360, -1.353745, -2.568015, -0.790628, 1.570796, 1.753156],accel_mss,speed_ms,0,blend_radius_m)
  movel([0.181837, -1.353098, -2.568452, -0.790839, 1.570796, 1.752633],accel_mss,speed_ms,0,blend_radius_m)
  movel([0.183063, -1.352762, -2.568679, -0.790948, 1.570796, 1.753859],accel_mss,speed_ms,0,blend_radius_m)
  movel([0.183512, -1.352645, -2.568758, -0.790987, 1.570796, 1.754308],accel_mss,speed_ms,0,blend_radius_m)
  movel([0.183955, -1.352542, -2.568827, -0.791020, 1.570796, 1.754752],accel_mss,speed_ms,0,blend_radius_m)
  movel([0.188162, -1.351613, -2.569452, -0.791324, 1.570796, 1.758958],accel_mss,speed_ms,0,blend_radius_m)
  movel([0.193088, -1.350554, -2.570163, -0.791672, 1.570796, 1.763885],accel_mss,speed_ms,0,blend_radius_m)
  movel([0.198699, -1.349384, -2.570947, -0.792058, 1.570796, 1.769495],accel_mss,speed_ms,0,blend_radius_m)
  movel([0.213116, -1.346499, -2.572872, -0.793018, 1.570796, 1.783912],accel_mss,speed_ms,0,blend_radius_m)
  movel([0.212938, -1.347258, -2.572367, -0.792765, 1.570796, 1.783735],accel_mss,speed_ms,0,blend_radius_m)
  movel([0.212761, -1.348015, -2.571862, -0.792512, 1.570796, 1.783557],accel_mss,speed_ms,0,blend_radius_m)
  movel([0.213243, -1.348125, -2.571788, -0.792475, 1.570796, 1.784040],accel_mss,speed_ms,0,blend_radius_m)
  movel([0.215483, -1.348602, -2.571470, -0.792317, 1.570796, 1.786280],accel_mss,speed_ms,0,blend_radius_m)
